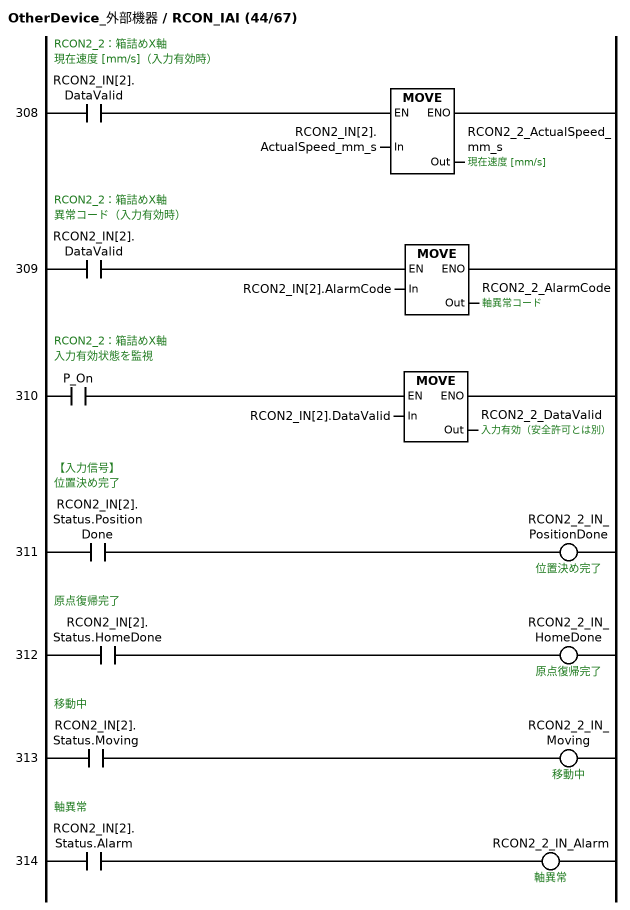
(* [picture p120: OtherDevice_外部機器 / RCON_IAI, rungs 308-314] *)
(* Rung 308: RCON2_2：箱詰めX軸 / 現在速度 [mm/s]（入力有効時） *)
IF RCON2_IN[2].DataValid THEN RCON2_2_ActualSpeed_mm_s := RCON2_IN[2].ActualSpeed_mm_s; END_IF;
(* Rung 309: RCON2_2：箱詰めX軸 / 異常コード（入力有効時） *)
IF RCON2_IN[2].DataValid THEN RCON2_2_AlarmCode := RCON2_IN[2].AlarmCode; END_IF;
(* Rung 310: RCON2_2：箱詰めX軸 / 入力有効状態を監視 *)
IF P_On THEN RCON2_2_DataValid := RCON2_IN[2].DataValid; END_IF;
(* Rung 311: 【入力信号】 / 位置決め完了 *)
RCON2_2_IN_PositionDone := RCON2_IN[2].Status.PositionDone;
(* Rung 312: 原点復帰完了 *)
RCON2_2_IN_HomeDone := RCON2_IN[2].Status.HomeDone;
(* Rung 313: 移動中 *)
RCON2_2_IN_Moving := RCON2_IN[2].Status.Moving;
(* Rung 314: 軸異常 *)
RCON2_2_IN_Alarm := RCON2_IN[2].Status.Alarm;

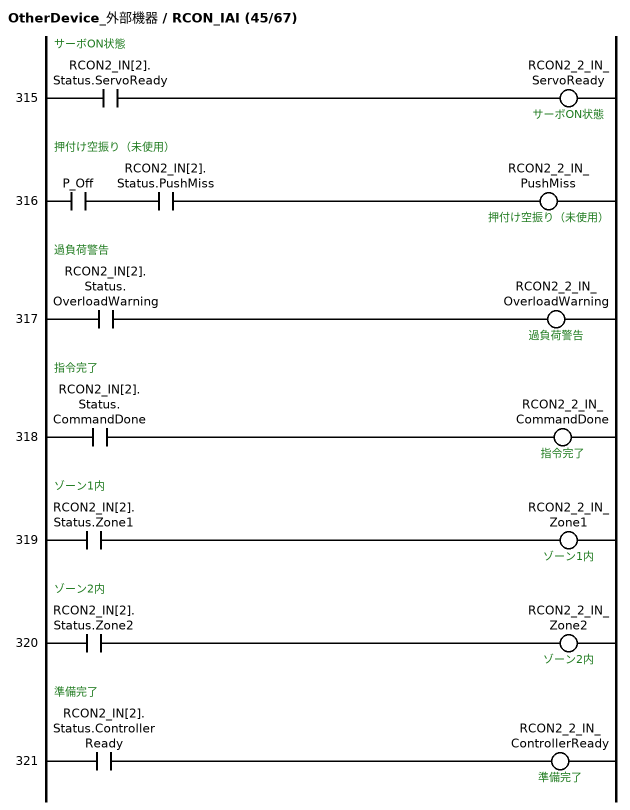
(* Rung 315: サーボON状態 *)
RCON2_2_IN_ServoReady := RCON2_IN[2].Status.ServoReady;
(* Rung 316: 押付け空振り（未使用） *)
RCON2_2_IN_PushMiss := P_Off AND RCON2_IN[2].Status.PushMiss;
(* Rung 317: 過負荷警告 *)
RCON2_2_IN_OverloadWarning := RCON2_IN[2].Status.OverloadWarning;
(* Rung 318: 指令完了 *)
RCON2_2_IN_CommandDone := RCON2_IN[2].Status.CommandDone;
(* Rung 319: ゾーン1内 *)
RCON2_2_IN_Zone1 := RCON2_IN[2].Status.Zone1;
(* Rung 320: ゾーン2内 *)
RCON2_2_IN_Zone2 := RCON2_IN[2].Status.Zone2;
(* Rung 321: 準備完了 *)
RCON2_2_IN_ControllerReady := RCON2_IN[2].Status.ControllerReady;

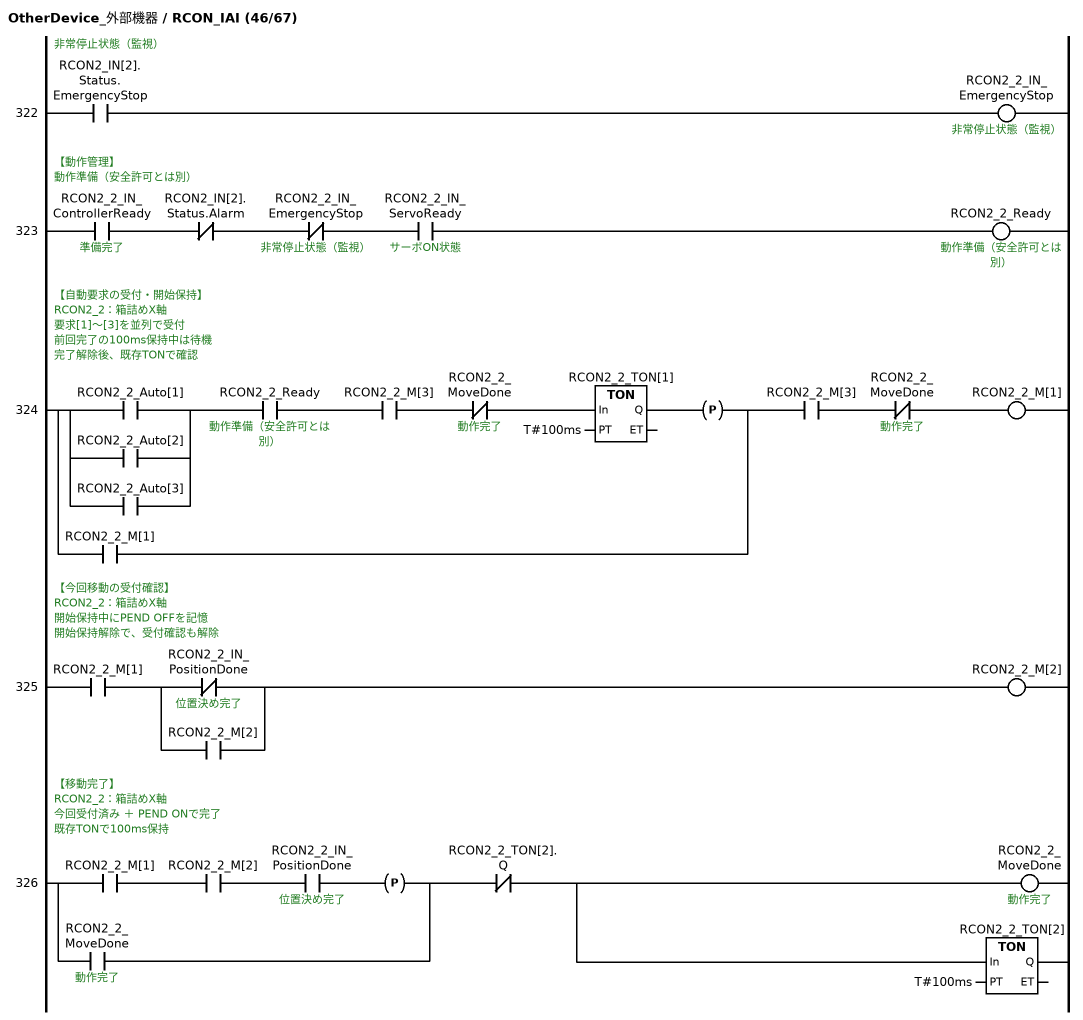
(* Rung 322: 非常停止状態（監視） *)
RCON2_2_IN_EmergencyStop := RCON2_IN[2].Status.EmergencyStop;
(* Rung 323: 【動作管理】 / 動作準備（安全許可とは別） *)
RCON2_2_Ready := RCON2_2_IN_ControllerReady AND NOT RCON2_IN[2].Status.Alarm AND NOT RCON2_2_IN_EmergencyStop AND RCON2_2_IN_ServoReady;
(* Rung 324: 【自動要求の受付・開始保持】 / RCON2_2：箱詰めX軸 / 要求[1]～[3]を並列で受付 / 前回完了の100ms保持中は待機 / 完了解除後、既存TONで確認 *)
RCON2_2_TON[1](In := (RCON2_2_Auto[1] OR RCON2_2_Auto[2] OR RCON2_2_Auto[3]) AND RCON2_2_Ready AND RCON2_2_M[3] AND NOT RCON2_2_MoveDone, PT := T#100ms);
_e30(CLK := RCON2_2_TON[1].Q);
RCON2_2_M[1] := (_e30.Q OR RCON2_2_M[1]) AND RCON2_2_M[3] AND NOT RCON2_2_MoveDone;
(* Rung 325: 【今回移動の受付確認】 / RCON2_2：箱詰めX軸 / 開始保持中にPEND OFFを記憶 / 開始保持解除で、受付確認も解除 *)
RCON2_2_M[2] := RCON2_2_M[1] AND (NOT RCON2_2_IN_PositionDone OR RCON2_2_M[2]);
(* Rung 326: 【移動完了】 / RCON2_2：箱詰めX軸 / 今回受付済み ＋ PEND ONで完了 / 既存TONで100ms保持 *)
_e31(CLK := RCON2_2_M[1] AND RCON2_2_M[2] AND RCON2_2_IN_PositionDone);
_p32 := (_e31.Q OR RCON2_2_MoveDone) AND NOT RCON2_2_TON[2].Q;
RCON2_2_MoveDone := _p32;
RCON2_2_TON[2](In := _p32, PT := T#100ms);

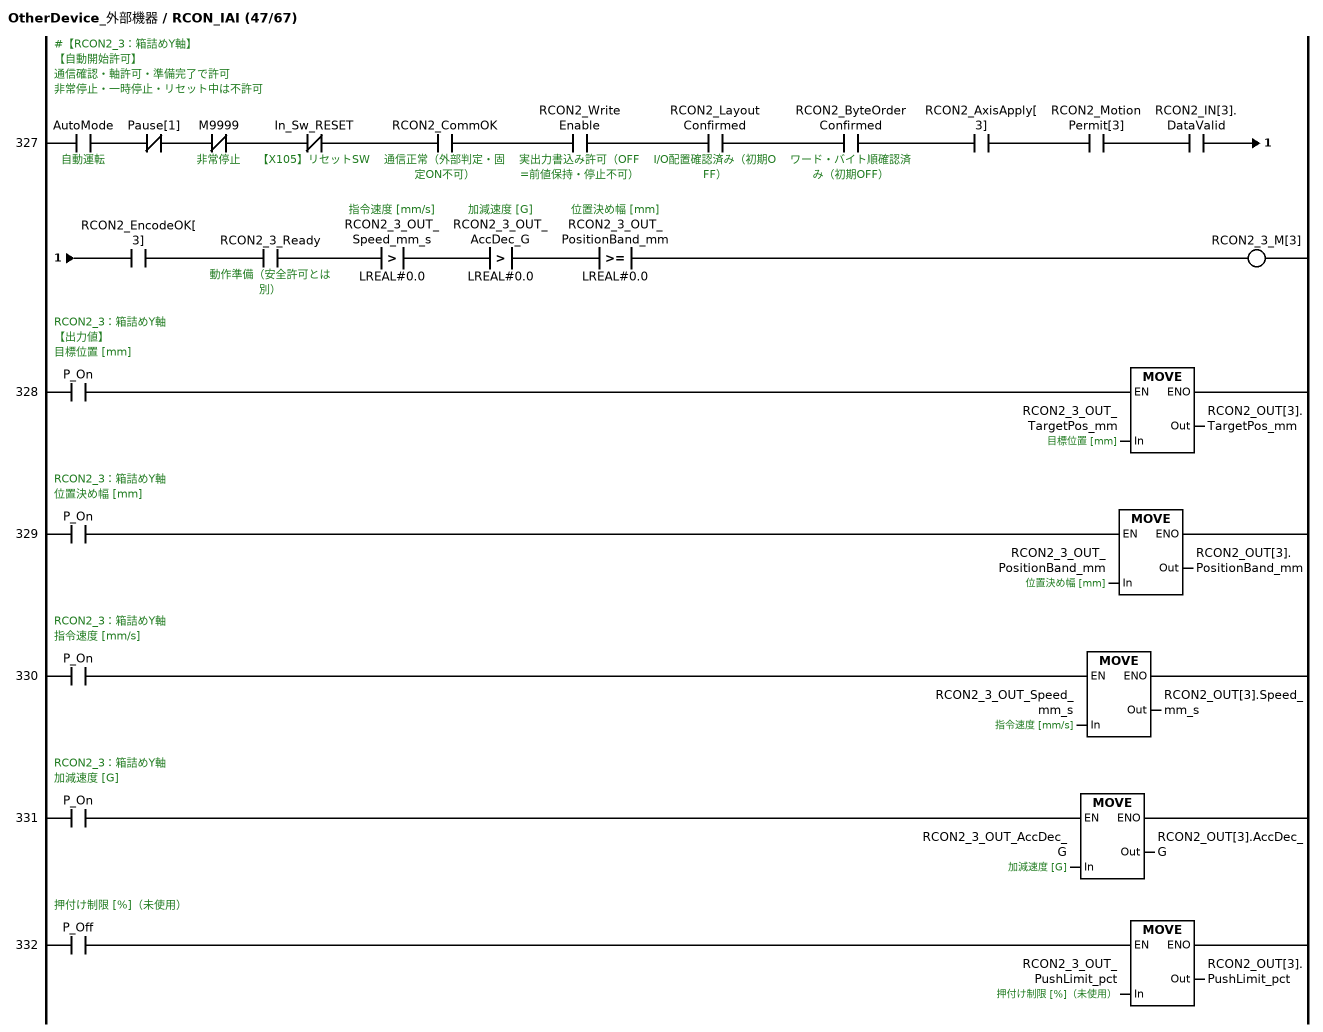
(* Rung 327: #【RCON2_3：箱詰めY軸】 / 【自動開始許可】 / 通信確認・軸許可・準備完了で許可 / 非常停止・一時停止・リセット中は不許可 *)
RCON2_3_M[3] := AutoMode AND NOT Pause[1] AND NOT M9999 AND NOT In_Sw_RESET AND RCON2_CommOK AND RCON2_WriteEnable AND RCON2_LayoutConfirmed AND RCON2_ByteOrderConfirmed AND RCON2_AxisApply[3] AND RCON2_MotionPermit[3] AND RCON2_IN[3].DataValid AND RCON2_EncodeOK[3] AND RCON2_3_Ready AND (RCON2_3_OUT_Speed_mm_s > LREAL#0.0) AND (RCON2_3_OUT_AccDec_G > LREAL#0.0) AND (RCON2_3_OUT_PositionBand_mm >= LREAL#0.0);
(* Rung 328: RCON2_3：箱詰めY軸 / 【出力値】 / 目標位置 [mm] *)
IF P_On THEN RCON2_OUT[3].TargetPos_mm := RCON2_3_OUT_TargetPos_mm; END_IF;
(* Rung 329: RCON2_3：箱詰めY軸 / 位置決め幅 [mm] *)
IF P_On THEN RCON2_OUT[3].PositionBand_mm := RCON2_3_OUT_PositionBand_mm; END_IF;
(* Rung 330: RCON2_3：箱詰めY軸 / 指令速度 [mm/s] *)
IF P_On THEN RCON2_OUT[3].Speed_mm_s := RCON2_3_OUT_Speed_mm_s; END_IF;
(* Rung 331: RCON2_3：箱詰めY軸 / 加減速度 [G] *)
IF P_On THEN RCON2_OUT[3].AccDec_G := RCON2_3_OUT_AccDec_G; END_IF;
(* Rung 332: 押付け制限 [%]（未使用） *)
IF P_Off THEN RCON2_OUT[3].PushLimit_pct := RCON2_3_OUT_PushLimit_pct; END_IF;

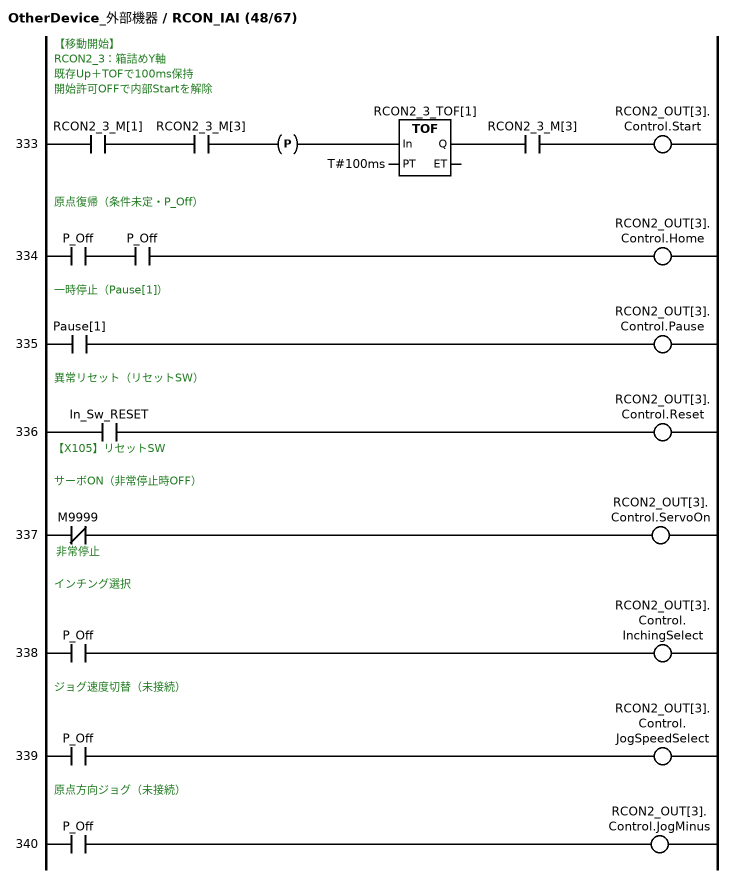
(* Rung 333: 【移動開始】 / RCON2_3：箱詰めY軸 / 既存Up＋TOFで100ms保持 / 開始許可OFFで内部Startを解除 *)
_e33(CLK := RCON2_3_M[1] AND RCON2_3_M[3]);
RCON2_3_TOF[1](In := _e33.Q, PT := T#100ms);
RCON2_OUT[3].Control.Start := RCON2_3_TOF[1].Q AND RCON2_3_M[3];
(* Rung 334: 原点復帰（条件未定・P_Off） *)
RCON2_OUT[3].Control.Home := P_Off AND P_Off;
(* Rung 335: 一時停止（Pause[1]） *)
RCON2_OUT[3].Control.Pause := Pause[1];
(* Rung 336: 異常リセット（リセットSW） *)
RCON2_OUT[3].Control.Reset := In_Sw_RESET;
(* Rung 337: サーボON（非常停止時OFF） *)
RCON2_OUT[3].Control.ServoOn := NOT M9999;
(* Rung 338: インチング選択 *)
RCON2_OUT[3].Control.InchingSelect := P_Off;
(* Rung 339: ジョグ速度切替（未接続） *)
RCON2_OUT[3].Control.JogSpeedSelect := P_Off;
(* Rung 340: 原点方向ジョグ（未接続） *)
RCON2_OUT[3].Control.JogMinus := P_Off;

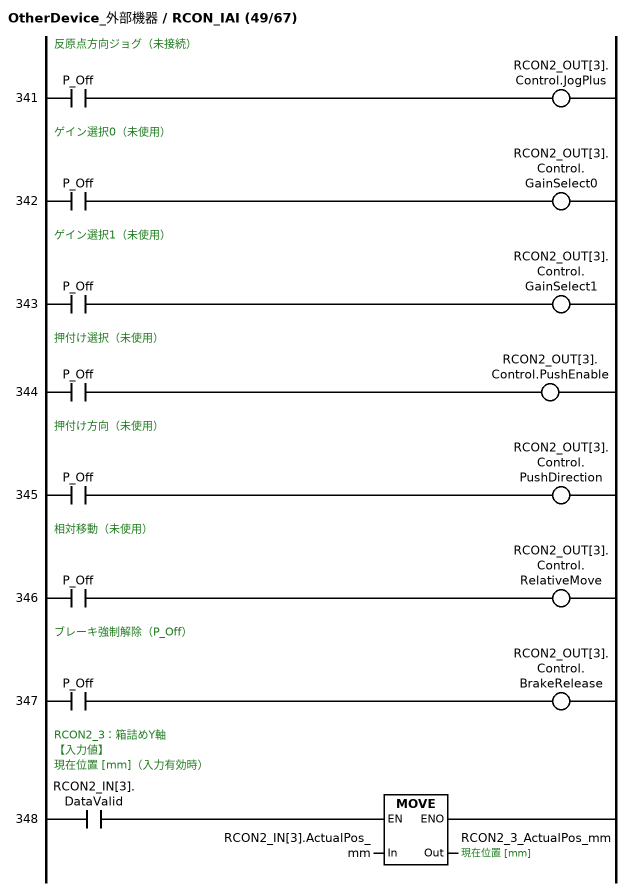
(* Rung 341: 反原点方向ジョグ（未接続） *)
RCON2_OUT[3].Control.JogPlus := P_Off;
(* Rung 342: ゲイン選択0（未使用） *)
RCON2_OUT[3].Control.GainSelect0 := P_Off;
(* Rung 343: ゲイン選択1（未使用） *)
RCON2_OUT[3].Control.GainSelect1 := P_Off;
(* Rung 344: 押付け選択（未使用） *)
RCON2_OUT[3].Control.PushEnable := P_Off;
(* Rung 345: 押付け方向（未使用） *)
RCON2_OUT[3].Control.PushDirection := P_Off;
(* Rung 346: 相対移動（未使用） *)
RCON2_OUT[3].Control.RelativeMove := P_Off;
(* Rung 347: ブレーキ強制解除（P_Off） *)
RCON2_OUT[3].Control.BrakeRelease := P_Off;
(* Rung 348: RCON2_3：箱詰めY軸 / 【入力値】 / 現在位置 [mm]（入力有効時） *)
IF RCON2_IN[3].DataValid THEN RCON2_3_ActualPos_mm := RCON2_IN[3].ActualPos_mm; END_IF;

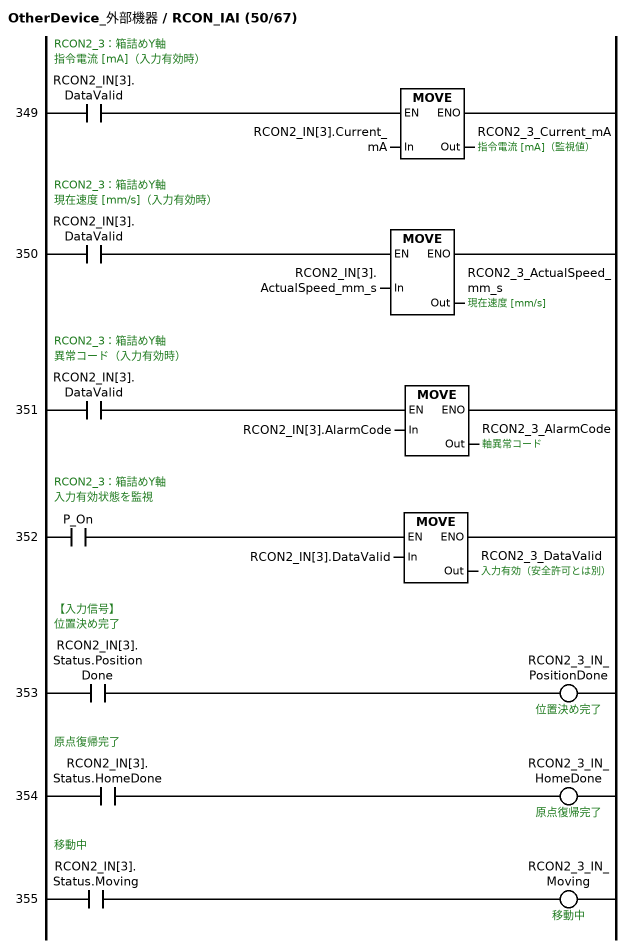
(* Rung 349: RCON2_3：箱詰めY軸 / 指令電流 [mA]（入力有効時） *)
IF RCON2_IN[3].DataValid THEN RCON2_3_Current_mA := RCON2_IN[3].Current_mA; END_IF;
(* Rung 350: RCON2_3：箱詰めY軸 / 現在速度 [mm/s]（入力有効時） *)
IF RCON2_IN[3].DataValid THEN RCON2_3_ActualSpeed_mm_s := RCON2_IN[3].ActualSpeed_mm_s; END_IF;
(* Rung 351: RCON2_3：箱詰めY軸 / 異常コード（入力有効時） *)
IF RCON2_IN[3].DataValid THEN RCON2_3_AlarmCode := RCON2_IN[3].AlarmCode; END_IF;
(* Rung 352: RCON2_3：箱詰めY軸 / 入力有効状態を監視 *)
IF P_On THEN RCON2_3_DataValid := RCON2_IN[3].DataValid; END_IF;
(* Rung 353: 【入力信号】 / 位置決め完了 *)
RCON2_3_IN_PositionDone := RCON2_IN[3].Status.PositionDone;
(* Rung 354: 原点復帰完了 *)
RCON2_3_IN_HomeDone := RCON2_IN[3].Status.HomeDone;
(* Rung 355: 移動中 *)
RCON2_3_IN_Moving := RCON2_IN[3].Status.Moving;

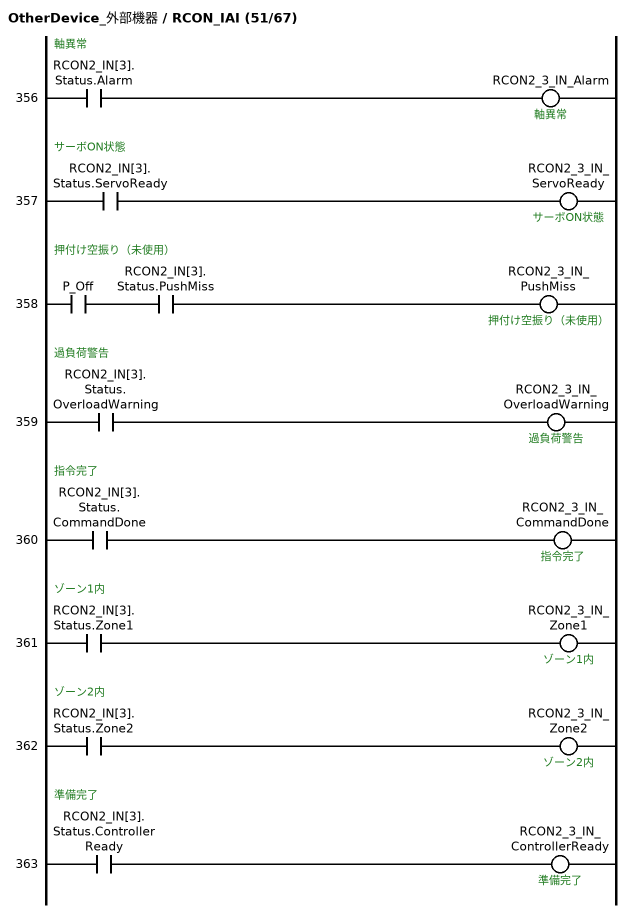
(* Rung 356: 軸異常 *)
RCON2_3_IN_Alarm := RCON2_IN[3].Status.Alarm;
(* Rung 357: サーボON状態 *)
RCON2_3_IN_ServoReady := RCON2_IN[3].Status.ServoReady;
(* Rung 358: 押付け空振り（未使用） *)
RCON2_3_IN_PushMiss := P_Off AND RCON2_IN[3].Status.PushMiss;
(* Rung 359: 過負荷警告 *)
RCON2_3_IN_OverloadWarning := RCON2_IN[3].Status.OverloadWarning;
(* Rung 360: 指令完了 *)
RCON2_3_IN_CommandDone := RCON2_IN[3].Status.CommandDone;
(* Rung 361: ゾーン1内 *)
RCON2_3_IN_Zone1 := RCON2_IN[3].Status.Zone1;
(* Rung 362: ゾーン2内 *)
RCON2_3_IN_Zone2 := RCON2_IN[3].Status.Zone2;
(* Rung 363: 準備完了 *)
RCON2_3_IN_ControllerReady := RCON2_IN[3].Status.ControllerReady;

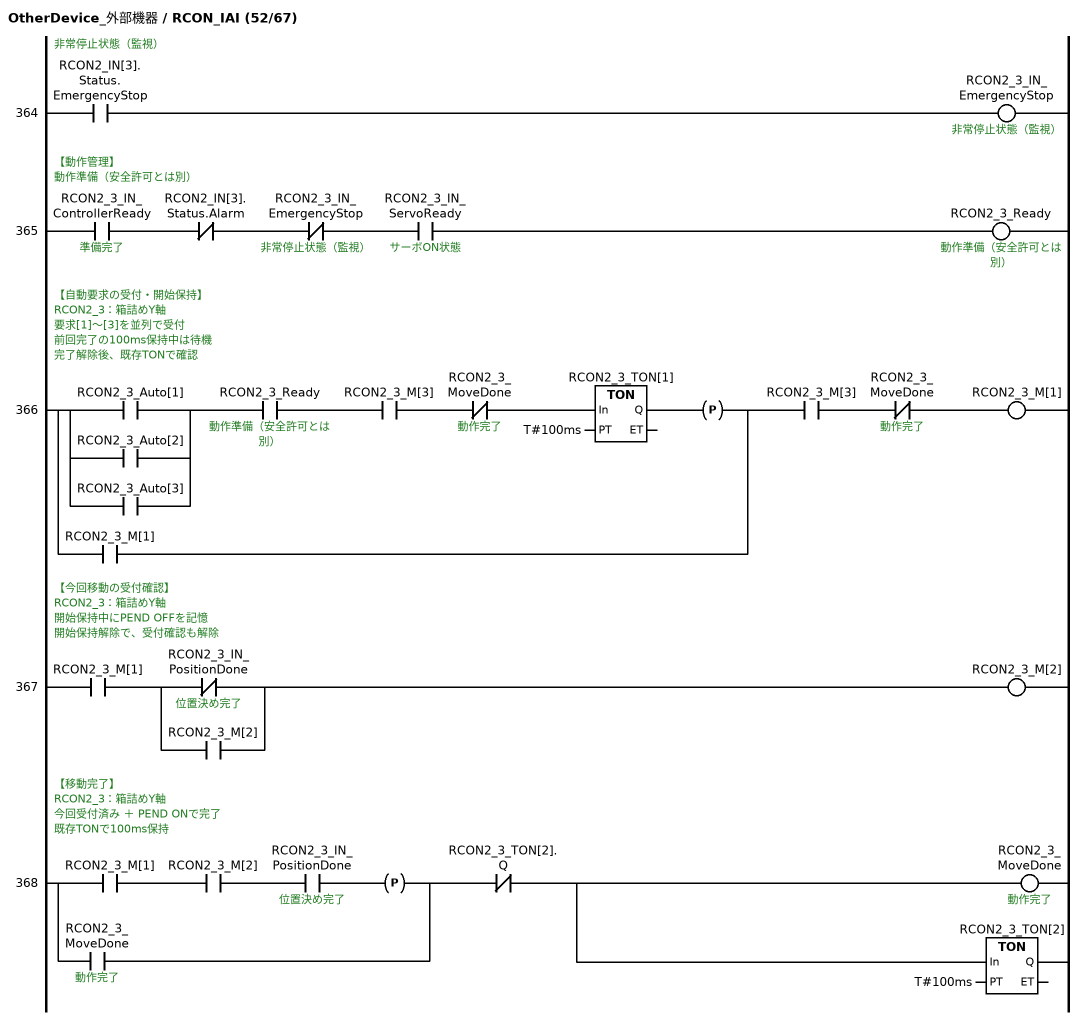
(* Rung 364: 非常停止状態（監視） *)
RCON2_3_IN_EmergencyStop := RCON2_IN[3].Status.EmergencyStop;
(* Rung 365: 【動作管理】 / 動作準備（安全許可とは別） *)
RCON2_3_Ready := RCON2_3_IN_ControllerReady AND NOT RCON2_IN[3].Status.Alarm AND NOT RCON2_3_IN_EmergencyStop AND RCON2_3_IN_ServoReady;
(* Rung 366: 【自動要求の受付・開始保持】 / RCON2_3：箱詰めY軸 / 要求[1]～[3]を並列で受付 / 前回完了の100ms保持中は待機 / 完了解除後、既存TONで確認 *)
RCON2_3_TON[1](In := (RCON2_3_Auto[1] OR RCON2_3_Auto[2] OR RCON2_3_Auto[3]) AND RCON2_3_Ready AND RCON2_3_M[3] AND NOT RCON2_3_MoveDone, PT := T#100ms);
_e34(CLK := RCON2_3_TON[1].Q);
RCON2_3_M[1] := (_e34.Q OR RCON2_3_M[1]) AND RCON2_3_M[3] AND NOT RCON2_3_MoveDone;
(* Rung 367: 【今回移動の受付確認】 / RCON2_3：箱詰めY軸 / 開始保持中にPEND OFFを記憶 / 開始保持解除で、受付確認も解除 *)
RCON2_3_M[2] := RCON2_3_M[1] AND (NOT RCON2_3_IN_PositionDone OR RCON2_3_M[2]);
(* Rung 368: 【移動完了】 / RCON2_3：箱詰めY軸 / 今回受付済み ＋ PEND ONで完了 / 既存TONで100ms保持 *)
_e35(CLK := RCON2_3_M[1] AND RCON2_3_M[2] AND RCON2_3_IN_PositionDone);
_p36 := (_e35.Q OR RCON2_3_MoveDone) AND NOT RCON2_3_TON[2].Q;
RCON2_3_MoveDone := _p36;
RCON2_3_TON[2](In := _p36, PT := T#100ms);

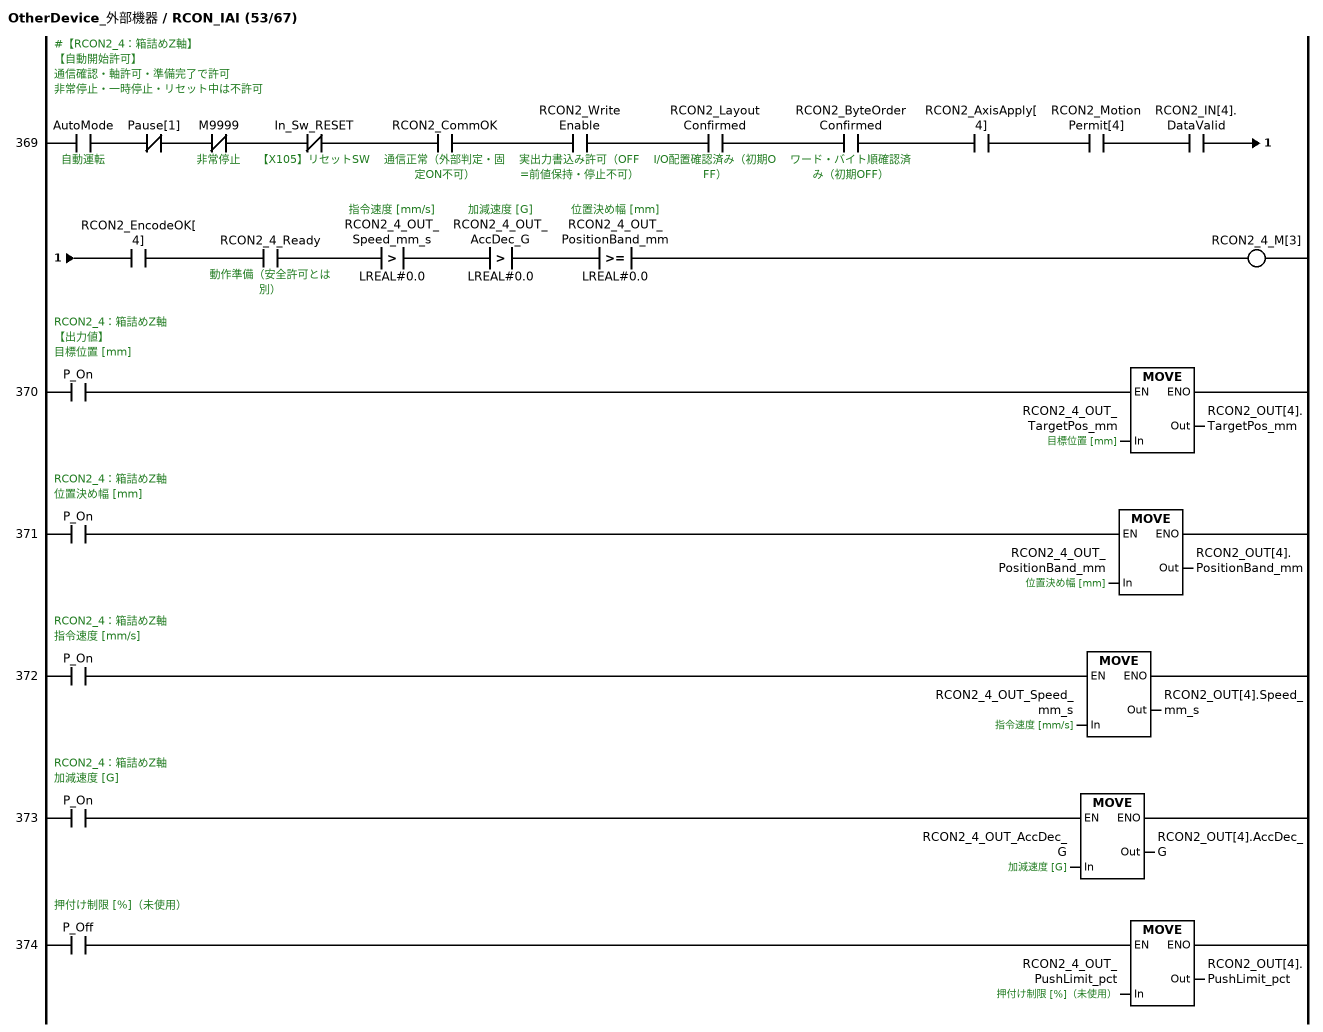
(* Rung 369: #【RCON2_4：箱詰めZ軸】 / 【自動開始許可】 / 通信確認・軸許可・準備完了で許可 / 非常停止・一時停止・リセット中は不許可 *)
RCON2_4_M[3] := AutoMode AND NOT Pause[1] AND NOT M9999 AND NOT In_Sw_RESET AND RCON2_CommOK AND RCON2_WriteEnable AND RCON2_LayoutConfirmed AND RCON2_ByteOrderConfirmed AND RCON2_AxisApply[4] AND RCON2_MotionPermit[4] AND RCON2_IN[4].DataValid AND RCON2_EncodeOK[4] AND RCON2_4_Ready AND (RCON2_4_OUT_Speed_mm_s > LREAL#0.0) AND (RCON2_4_OUT_AccDec_G > LREAL#0.0) AND (RCON2_4_OUT_PositionBand_mm >= LREAL#0.0);
(* Rung 370: RCON2_4：箱詰めZ軸 / 【出力値】 / 目標位置 [mm] *)
IF P_On THEN RCON2_OUT[4].TargetPos_mm := RCON2_4_OUT_TargetPos_mm; END_IF;
(* Rung 371: RCON2_4：箱詰めZ軸 / 位置決め幅 [mm] *)
IF P_On THEN RCON2_OUT[4].PositionBand_mm := RCON2_4_OUT_PositionBand_mm; END_IF;
(* Rung 372: RCON2_4：箱詰めZ軸 / 指令速度 [mm/s] *)
IF P_On THEN RCON2_OUT[4].Speed_mm_s := RCON2_4_OUT_Speed_mm_s; END_IF;
(* Rung 373: RCON2_4：箱詰めZ軸 / 加減速度 [G] *)
IF P_On THEN RCON2_OUT[4].AccDec_G := RCON2_4_OUT_AccDec_G; END_IF;
(* Rung 374: 押付け制限 [%]（未使用） *)
IF P_Off THEN RCON2_OUT[4].PushLimit_pct := RCON2_4_OUT_PushLimit_pct; END_IF;

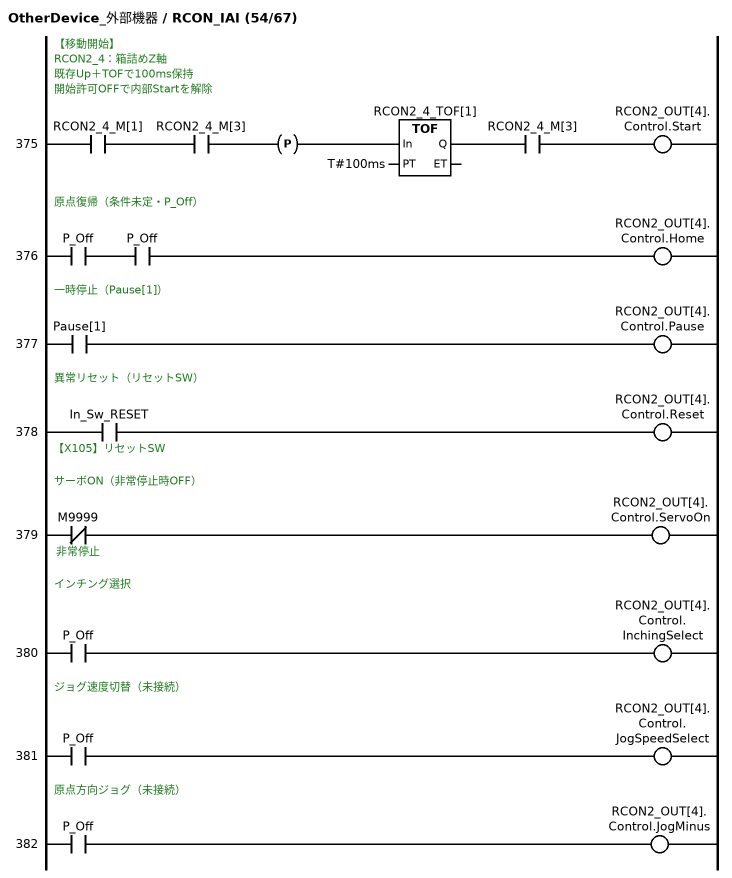
(* Rung 375: 【移動開始】 / RCON2_4：箱詰めZ軸 / 既存Up＋TOFで100ms保持 / 開始許可OFFで内部Startを解除 *)
_e37(CLK := RCON2_4_M[1] AND RCON2_4_M[3]);
RCON2_4_TOF[1](In := _e37.Q, PT := T#100ms);
RCON2_OUT[4].Control.Start := RCON2_4_TOF[1].Q AND RCON2_4_M[3];
(* Rung 376: 原点復帰（条件未定・P_Off） *)
RCON2_OUT[4].Control.Home := P_Off AND P_Off;
(* Rung 377: 一時停止（Pause[1]） *)
RCON2_OUT[4].Control.Pause := Pause[1];
(* Rung 378: 異常リセット（リセットSW） *)
RCON2_OUT[4].Control.Reset := In_Sw_RESET;
(* Rung 379: サーボON（非常停止時OFF） *)
RCON2_OUT[4].Control.ServoOn := NOT M9999;
(* Rung 380: インチング選択 *)
RCON2_OUT[4].Control.InchingSelect := P_Off;
(* Rung 381: ジョグ速度切替（未接続） *)
RCON2_OUT[4].Control.JogSpeedSelect := P_Off;
(* Rung 382: 原点方向ジョグ（未接続） *)
RCON2_OUT[4].Control.JogMinus := P_Off;

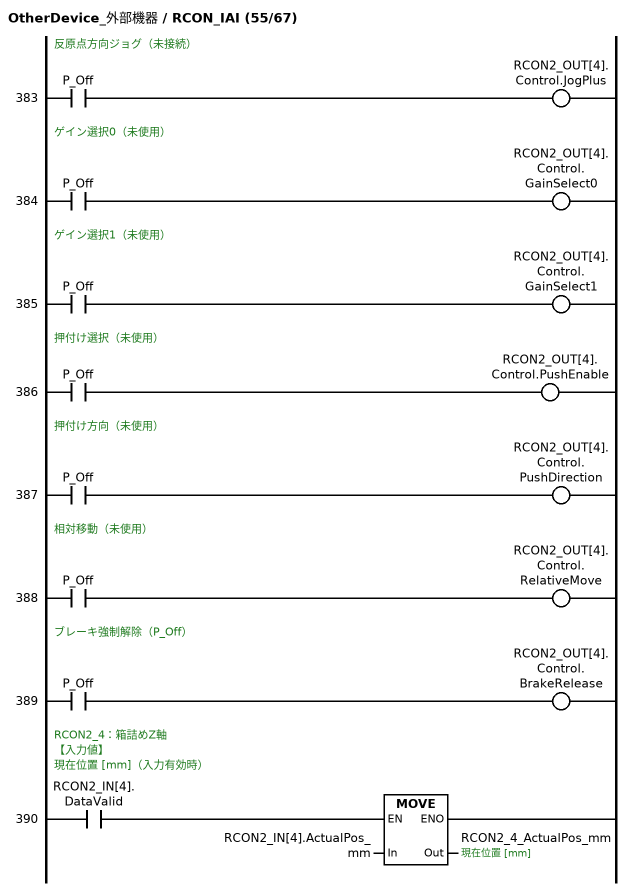
(* Rung 383: 反原点方向ジョグ（未接続） *)
RCON2_OUT[4].Control.JogPlus := P_Off;
(* Rung 384: ゲイン選択0（未使用） *)
RCON2_OUT[4].Control.GainSelect0 := P_Off;
(* Rung 385: ゲイン選択1（未使用） *)
RCON2_OUT[4].Control.GainSelect1 := P_Off;
(* Rung 386: 押付け選択（未使用） *)
RCON2_OUT[4].Control.PushEnable := P_Off;
(* Rung 387: 押付け方向（未使用） *)
RCON2_OUT[4].Control.PushDirection := P_Off;
(* Rung 388: 相対移動（未使用） *)
RCON2_OUT[4].Control.RelativeMove := P_Off;
(* Rung 389: ブレーキ強制解除（P_Off） *)
RCON2_OUT[4].Control.BrakeRelease := P_Off;
(* Rung 390: RCON2_4：箱詰めZ軸 / 【入力値】 / 現在位置 [mm]（入力有効時） *)
IF RCON2_IN[4].DataValid THEN RCON2_4_ActualPos_mm := RCON2_IN[4].ActualPos_mm; END_IF;

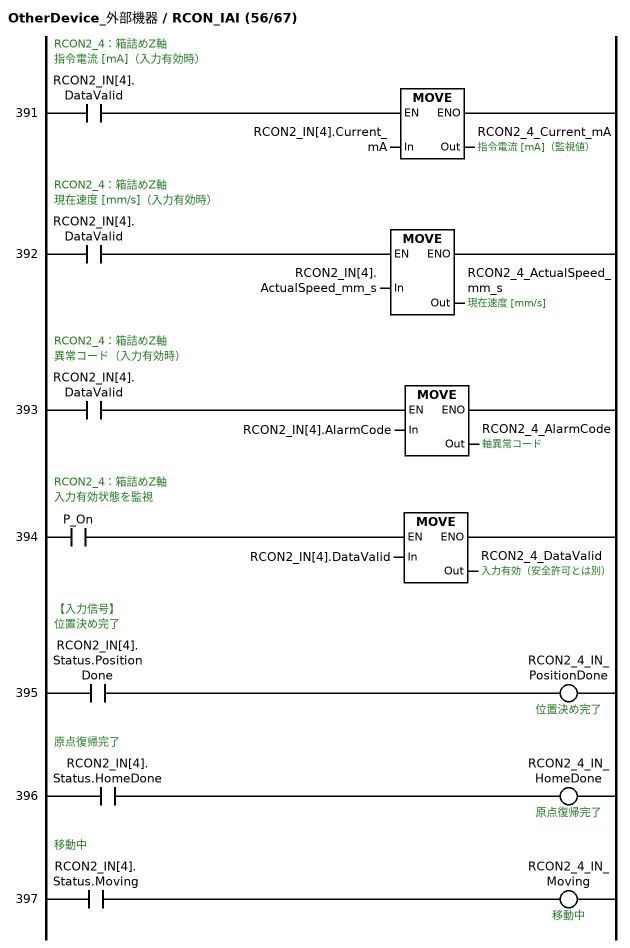
(* Rung 391: RCON2_4：箱詰めZ軸 / 指令電流 [mA]（入力有効時） *)
IF RCON2_IN[4].DataValid THEN RCON2_4_Current_mA := RCON2_IN[4].Current_mA; END_IF;
(* Rung 392: RCON2_4：箱詰めZ軸 / 現在速度 [mm/s]（入力有効時） *)
IF RCON2_IN[4].DataValid THEN RCON2_4_ActualSpeed_mm_s := RCON2_IN[4].ActualSpeed_mm_s; END_IF;
(* Rung 393: RCON2_4：箱詰めZ軸 / 異常コード（入力有効時） *)
IF RCON2_IN[4].DataValid THEN RCON2_4_AlarmCode := RCON2_IN[4].AlarmCode; END_IF;
(* Rung 394: RCON2_4：箱詰めZ軸 / 入力有効状態を監視 *)
IF P_On THEN RCON2_4_DataValid := RCON2_IN[4].DataValid; END_IF;
(* Rung 395: 【入力信号】 / 位置決め完了 *)
RCON2_4_IN_PositionDone := RCON2_IN[4].Status.PositionDone;
(* Rung 396: 原点復帰完了 *)
RCON2_4_IN_HomeDone := RCON2_IN[4].Status.HomeDone;
(* Rung 397: 移動中 *)
RCON2_4_IN_Moving := RCON2_IN[4].Status.Moving;

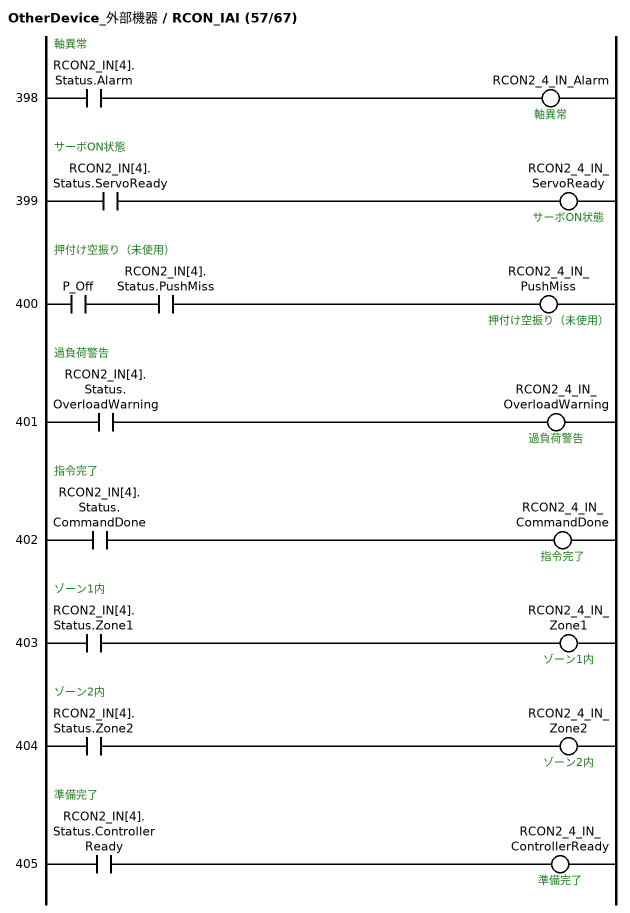
(* Rung 398: 軸異常 *)
RCON2_4_IN_Alarm := RCON2_IN[4].Status.Alarm;
(* Rung 399: サーボON状態 *)
RCON2_4_IN_ServoReady := RCON2_IN[4].Status.ServoReady;
(* Rung 400: 押付け空振り（未使用） *)
RCON2_4_IN_PushMiss := P_Off AND RCON2_IN[4].Status.PushMiss;
(* Rung 401: 過負荷警告 *)
RCON2_4_IN_OverloadWarning := RCON2_IN[4].Status.OverloadWarning;
(* Rung 402: 指令完了 *)
RCON2_4_IN_CommandDone := RCON2_IN[4].Status.CommandDone;
(* Rung 403: ゾーン1内 *)
RCON2_4_IN_Zone1 := RCON2_IN[4].Status.Zone1;
(* Rung 404: ゾーン2内 *)
RCON2_4_IN_Zone2 := RCON2_IN[4].Status.Zone2;
(* Rung 405: 準備完了 *)
RCON2_4_IN_ControllerReady := RCON2_IN[4].Status.ControllerReady;

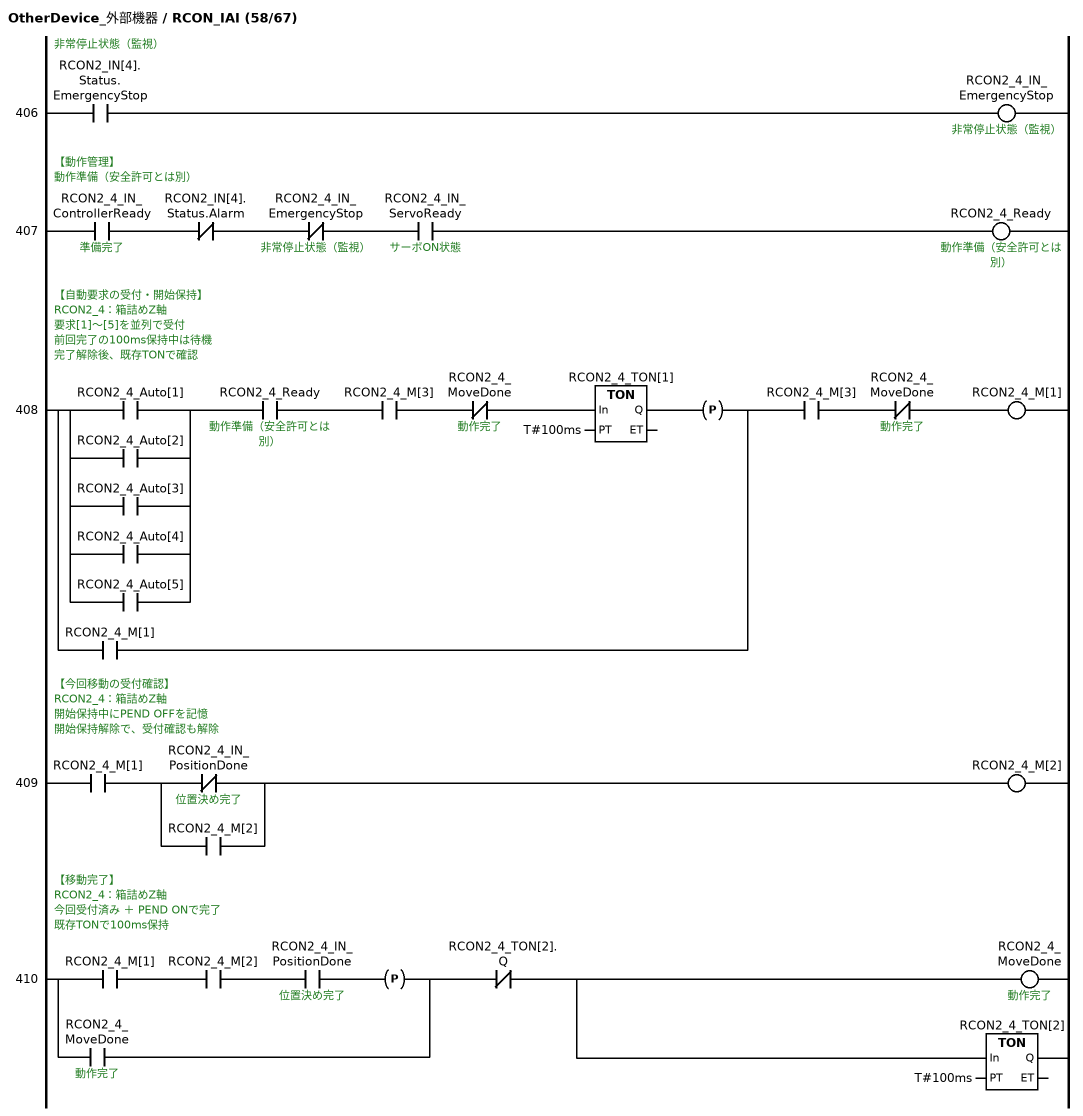
(* Rung 406: 非常停止状態（監視） *)
RCON2_4_IN_EmergencyStop := RCON2_IN[4].Status.EmergencyStop;
(* Rung 407: 【動作管理】 / 動作準備（安全許可とは別） *)
RCON2_4_Ready := RCON2_4_IN_ControllerReady AND NOT RCON2_IN[4].Status.Alarm AND NOT RCON2_4_IN_EmergencyStop AND RCON2_4_IN_ServoReady;
(* Rung 408: 【自動要求の受付・開始保持】 / RCON2_4：箱詰めZ軸 / 要求[1]～[5]を並列で受付 / 前回完了の100ms保持中は待機 / 完了解除後、既存TONで確認 *)
RCON2_4_TON[1](In := (RCON2_4_Auto[1] OR RCON2_4_Auto[2] OR RCON2_4_Auto[3] OR RCON2_4_Auto[4] OR RCON2_4_Auto[5]) AND RCON2_4_Ready AND RCON2_4_M[3] AND NOT RCON2_4_MoveDone, PT := T#100ms);
_e38(CLK := RCON2_4_TON[1].Q);
RCON2_4_M[1] := (_e38.Q OR RCON2_4_M[1]) AND RCON2_4_M[3] AND NOT RCON2_4_MoveDone;
(* Rung 409: 【今回移動の受付確認】 / RCON2_4：箱詰めZ軸 / 開始保持中にPEND OFFを記憶 / 開始保持解除で、受付確認も解除 *)
RCON2_4_M[2] := RCON2_4_M[1] AND (NOT RCON2_4_IN_PositionDone OR RCON2_4_M[2]);
(* Rung 410: 【移動完了】 / RCON2_4：箱詰めZ軸 / 今回受付済み ＋ PEND ONで完了 / 既存TONで100ms保持 *)
_e39(CLK := RCON2_4_M[1] AND RCON2_4_M[2] AND RCON2_4_IN_PositionDone);
_p40 := (_e39.Q OR RCON2_4_MoveDone) AND NOT RCON2_4_TON[2].Q;
RCON2_4_MoveDone := _p40;
RCON2_4_TON[2](In := _p40, PT := T#100ms);

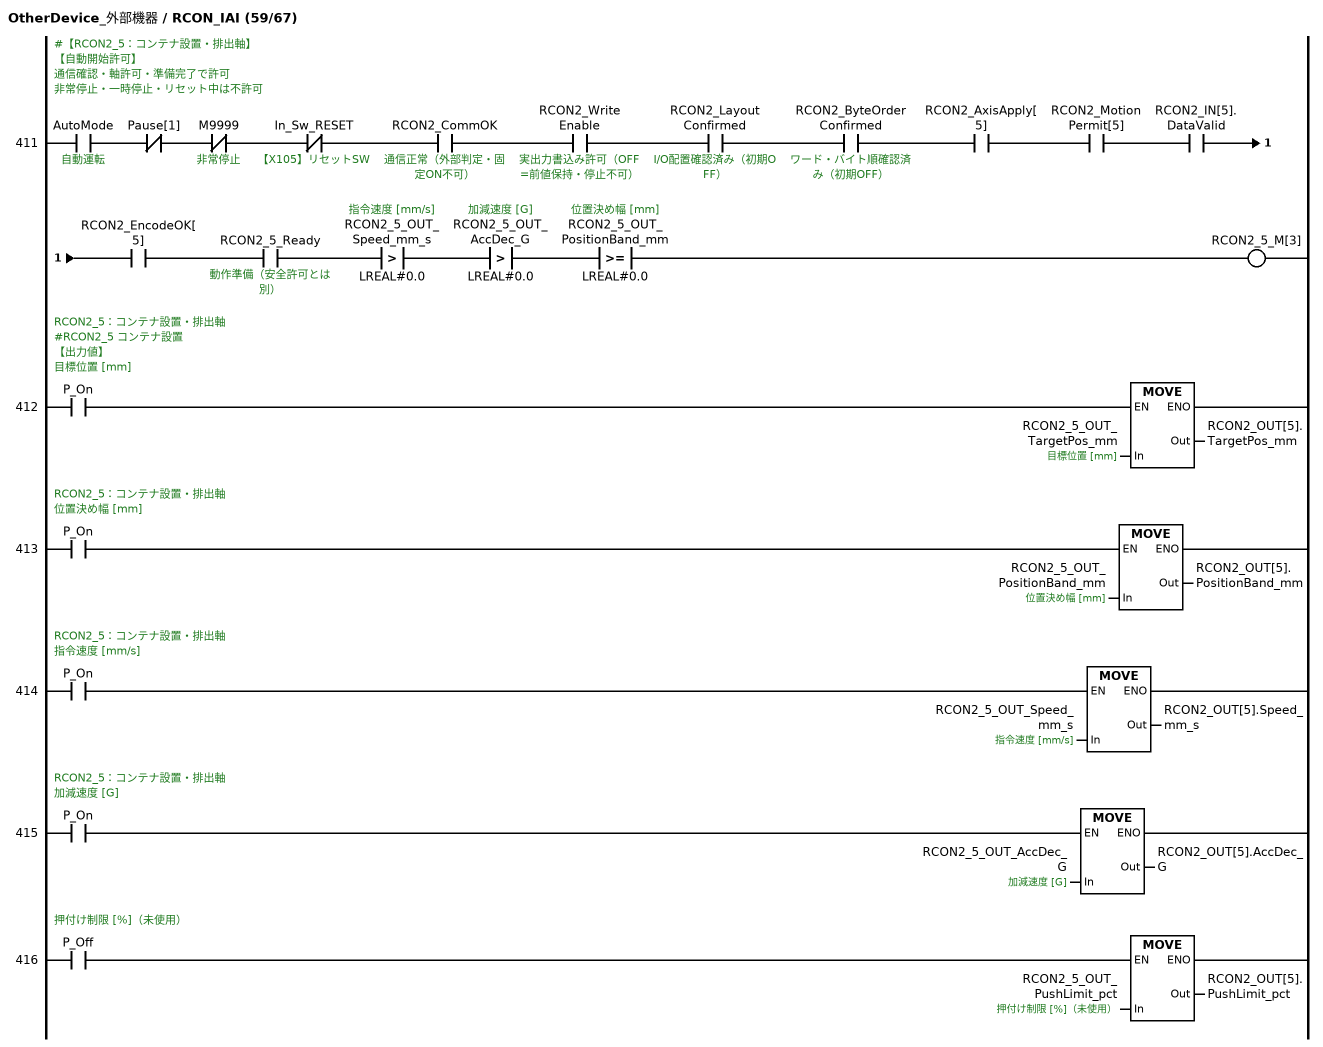
(* Rung 411: #【RCON2_5：コンテナ設置・排出軸】 / 【自動開始許可】 / 通信確認・軸許可・準備完了で許可 / 非常停止・一時停止・リセット中は不許可 *)
RCON2_5_M[3] := AutoMode AND NOT Pause[1] AND NOT M9999 AND NOT In_Sw_RESET AND RCON2_CommOK AND RCON2_WriteEnable AND RCON2_LayoutConfirmed AND RCON2_ByteOrderConfirmed AND RCON2_AxisApply[5] AND RCON2_MotionPermit[5] AND RCON2_IN[5].DataValid AND RCON2_EncodeOK[5] AND RCON2_5_Ready AND (RCON2_5_OUT_Speed_mm_s > LREAL#0.0) AND (RCON2_5_OUT_AccDec_G > LREAL#0.0) AND (RCON2_5_OUT_PositionBand_mm >= LREAL#0.0);
(* Rung 412: RCON2_5：コンテナ設置・排出軸 / #RCON2_5 コンテナ設置 / 【出力値】 / 目標位置 [mm] *)
IF P_On THEN RCON2_OUT[5].TargetPos_mm := RCON2_5_OUT_TargetPos_mm; END_IF;
(* Rung 413: RCON2_5：コンテナ設置・排出軸 / 位置決め幅 [mm] *)
IF P_On THEN RCON2_OUT[5].PositionBand_mm := RCON2_5_OUT_PositionBand_mm; END_IF;
(* Rung 414: RCON2_5：コンテナ設置・排出軸 / 指令速度 [mm/s] *)
IF P_On THEN RCON2_OUT[5].Speed_mm_s := RCON2_5_OUT_Speed_mm_s; END_IF;
(* Rung 415: RCON2_5：コンテナ設置・排出軸 / 加減速度 [G] *)
IF P_On THEN RCON2_OUT[5].AccDec_G := RCON2_5_OUT_AccDec_G; END_IF;
(* Rung 416: 押付け制限 [%]（未使用） *)
IF P_Off THEN RCON2_OUT[5].PushLimit_pct := RCON2_5_OUT_PushLimit_pct; END_IF;

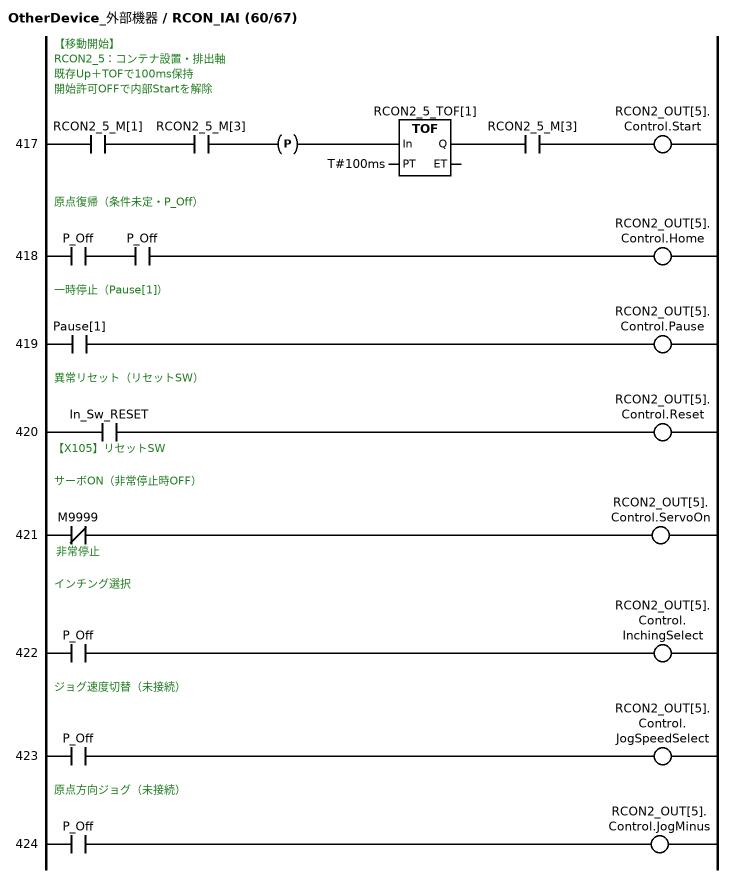
(* Rung 417: 【移動開始】 / RCON2_5：コンテナ設置・排出軸 / 既存Up＋TOFで100ms保持 / 開始許可OFFで内部Startを解除 *)
_e41(CLK := RCON2_5_M[1] AND RCON2_5_M[3]);
RCON2_5_TOF[1](In := _e41.Q, PT := T#100ms);
RCON2_OUT[5].Control.Start := RCON2_5_TOF[1].Q AND RCON2_5_M[3];
(* Rung 418: 原点復帰（条件未定・P_Off） *)
RCON2_OUT[5].Control.Home := P_Off AND P_Off;
(* Rung 419: 一時停止（Pause[1]） *)
RCON2_OUT[5].Control.Pause := Pause[1];
(* Rung 420: 異常リセット（リセットSW） *)
RCON2_OUT[5].Control.Reset := In_Sw_RESET;
(* Rung 421: サーボON（非常停止時OFF） *)
RCON2_OUT[5].Control.ServoOn := NOT M9999;
(* Rung 422: インチング選択 *)
RCON2_OUT[5].Control.InchingSelect := P_Off;
(* Rung 423: ジョグ速度切替（未接続） *)
RCON2_OUT[5].Control.JogSpeedSelect := P_Off;
(* Rung 424: 原点方向ジョグ（未接続） *)
RCON2_OUT[5].Control.JogMinus := P_Off;

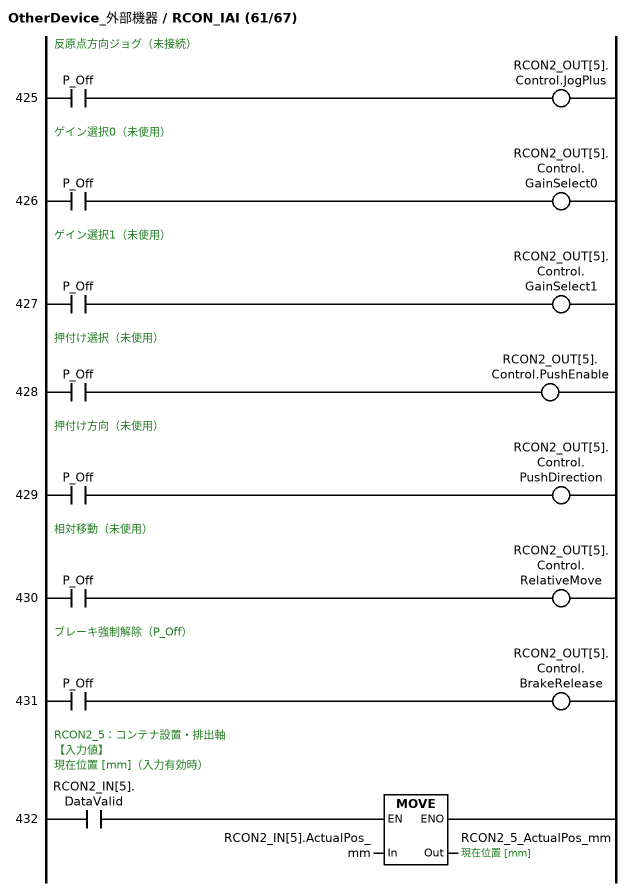
(* Rung 425: 反原点方向ジョグ（未接続） *)
RCON2_OUT[5].Control.JogPlus := P_Off;
(* Rung 426: ゲイン選択0（未使用） *)
RCON2_OUT[5].Control.GainSelect0 := P_Off;
(* Rung 427: ゲイン選択1（未使用） *)
RCON2_OUT[5].Control.GainSelect1 := P_Off;
(* Rung 428: 押付け選択（未使用） *)
RCON2_OUT[5].Control.PushEnable := P_Off;
(* Rung 429: 押付け方向（未使用） *)
RCON2_OUT[5].Control.PushDirection := P_Off;
(* Rung 430: 相対移動（未使用） *)
RCON2_OUT[5].Control.RelativeMove := P_Off;
(* Rung 431: ブレーキ強制解除（P_Off） *)
RCON2_OUT[5].Control.BrakeRelease := P_Off;
(* Rung 432: RCON2_5：コンテナ設置・排出軸 / 【入力値】 / 現在位置 [mm]（入力有効時） *)
IF RCON2_IN[5].DataValid THEN RCON2_5_ActualPos_mm := RCON2_IN[5].ActualPos_mm; END_IF;

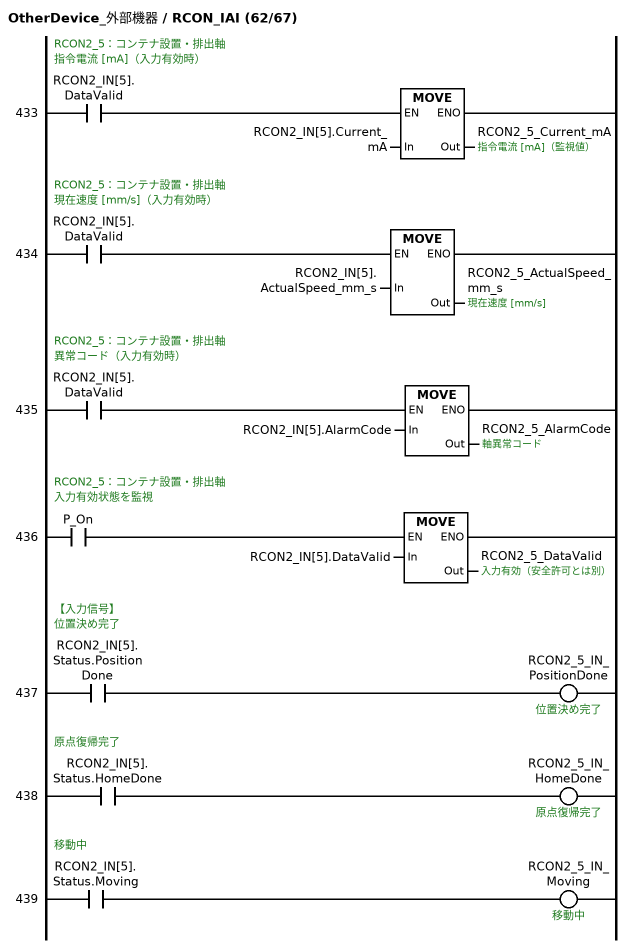
(* Rung 433: RCON2_5：コンテナ設置・排出軸 / 指令電流 [mA]（入力有効時） *)
IF RCON2_IN[5].DataValid THEN RCON2_5_Current_mA := RCON2_IN[5].Current_mA; END_IF;
(* Rung 434: RCON2_5：コンテナ設置・排出軸 / 現在速度 [mm/s]（入力有効時） *)
IF RCON2_IN[5].DataValid THEN RCON2_5_ActualSpeed_mm_s := RCON2_IN[5].ActualSpeed_mm_s; END_IF;
(* Rung 435: RCON2_5：コンテナ設置・排出軸 / 異常コード（入力有効時） *)
IF RCON2_IN[5].DataValid THEN RCON2_5_AlarmCode := RCON2_IN[5].AlarmCode; END_IF;
(* Rung 436: RCON2_5：コンテナ設置・排出軸 / 入力有効状態を監視 *)
IF P_On THEN RCON2_5_DataValid := RCON2_IN[5].DataValid; END_IF;
(* Rung 437: 【入力信号】 / 位置決め完了 *)
RCON2_5_IN_PositionDone := RCON2_IN[5].Status.PositionDone;
(* Rung 438: 原点復帰完了 *)
RCON2_5_IN_HomeDone := RCON2_IN[5].Status.HomeDone;
(* Rung 439: 移動中 *)
RCON2_5_IN_Moving := RCON2_IN[5].Status.Moving;

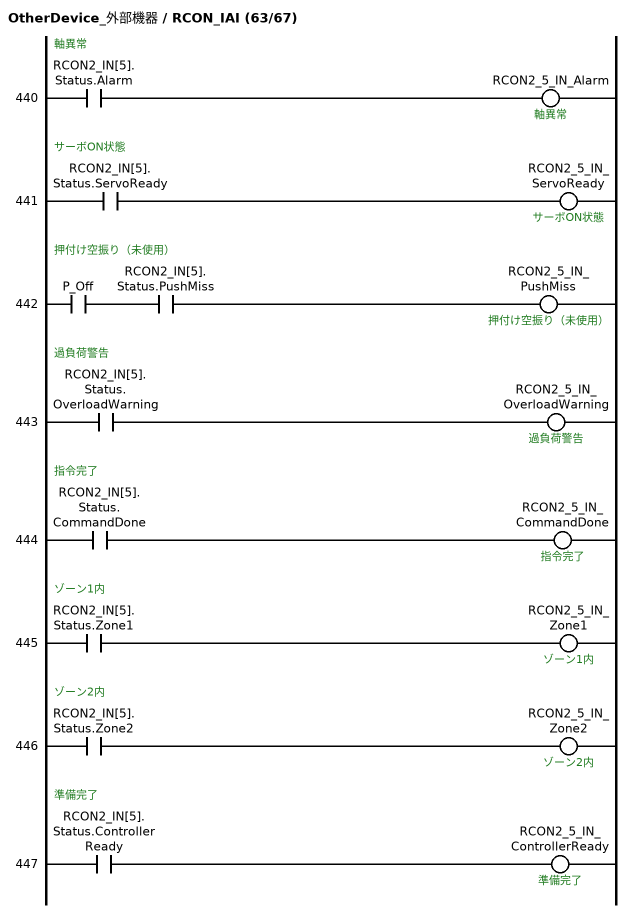
(* Rung 440: 軸異常 *)
RCON2_5_IN_Alarm := RCON2_IN[5].Status.Alarm;
(* Rung 441: サーボON状態 *)
RCON2_5_IN_ServoReady := RCON2_IN[5].Status.ServoReady;
(* Rung 442: 押付け空振り（未使用） *)
RCON2_5_IN_PushMiss := P_Off AND RCON2_IN[5].Status.PushMiss;
(* Rung 443: 過負荷警告 *)
RCON2_5_IN_OverloadWarning := RCON2_IN[5].Status.OverloadWarning;
(* Rung 444: 指令完了 *)
RCON2_5_IN_CommandDone := RCON2_IN[5].Status.CommandDone;
(* Rung 445: ゾーン1内 *)
RCON2_5_IN_Zone1 := RCON2_IN[5].Status.Zone1;
(* Rung 446: ゾーン2内 *)
RCON2_5_IN_Zone2 := RCON2_IN[5].Status.Zone2;
(* Rung 447: 準備完了 *)
RCON2_5_IN_ControllerReady := RCON2_IN[5].Status.ControllerReady;

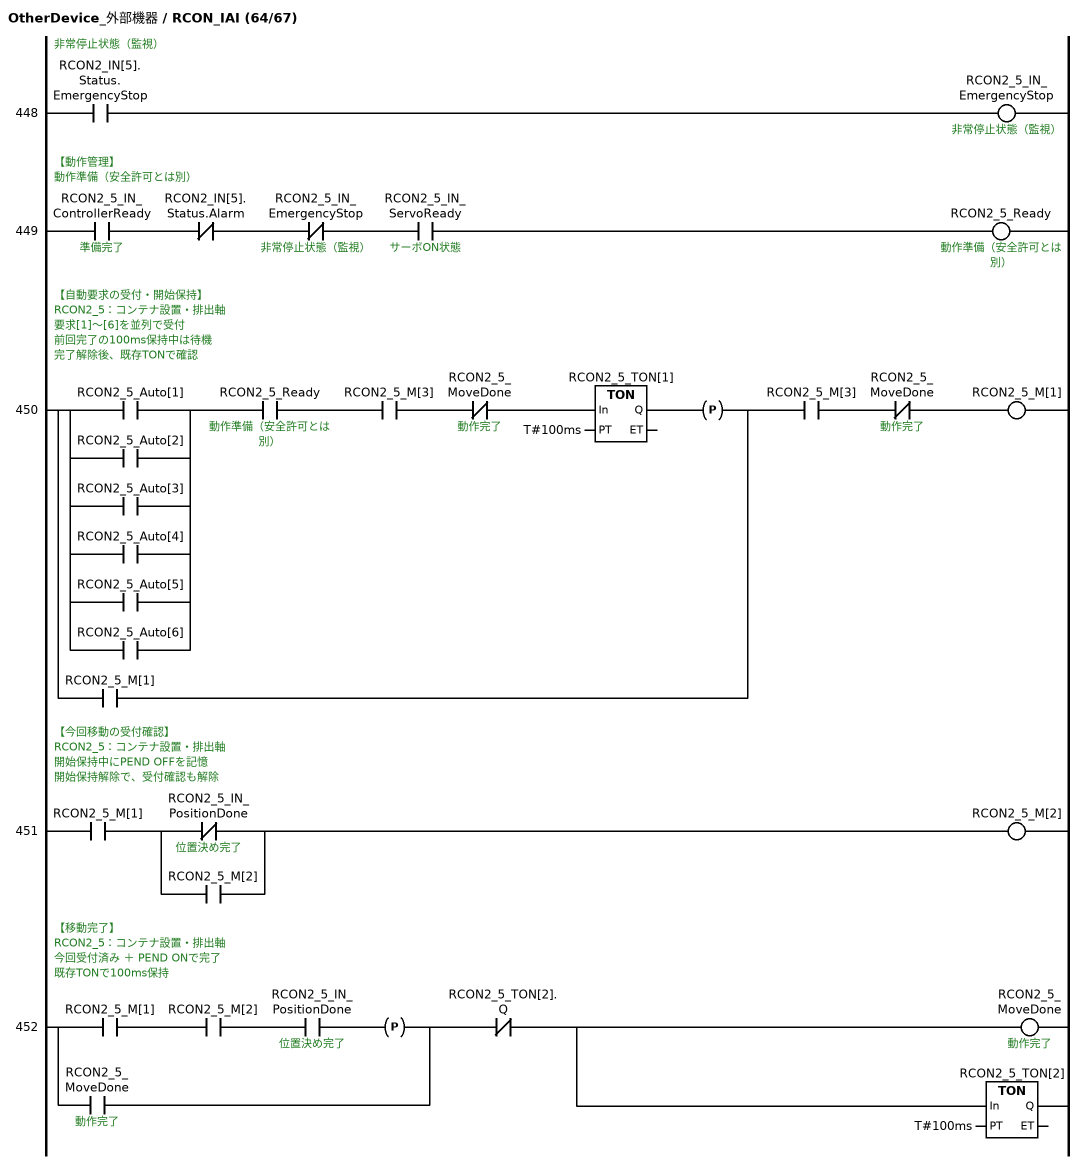
(* Rung 448: 非常停止状態（監視） *)
RCON2_5_IN_EmergencyStop := RCON2_IN[5].Status.EmergencyStop;
(* Rung 449: 【動作管理】 / 動作準備（安全許可とは別） *)
RCON2_5_Ready := RCON2_5_IN_ControllerReady AND NOT RCON2_IN[5].Status.Alarm AND NOT RCON2_5_IN_EmergencyStop AND RCON2_5_IN_ServoReady;
(* Rung 450: 【自動要求の受付・開始保持】 / RCON2_5：コンテナ設置・排出軸 / 要求[1]～[6]を並列で受付 / 前回完了の100ms保持中は待機 / 完了解除後、既存TONで確認 *)
RCON2_5_TON[1](In := (RCON2_5_Auto[1] OR RCON2_5_Auto[2] OR RCON2_5_Auto[3] OR RCON2_5_Auto[4] OR RCON2_5_Auto[5] OR RCON2_5_Auto[6]) AND RCON2_5_Ready AND RCON2_5_M[3] AND NOT RCON2_5_MoveDone, PT := T#100ms);
_e42(CLK := RCON2_5_TON[1].Q);
RCON2_5_M[1] := (_e42.Q OR RCON2_5_M[1]) AND RCON2_5_M[3] AND NOT RCON2_5_MoveDone;
(* Rung 451: 【今回移動の受付確認】 / RCON2_5：コンテナ設置・排出軸 / 開始保持中にPEND OFFを記憶 / 開始保持解除で、受付確認も解除 *)
RCON2_5_M[2] := RCON2_5_M[1] AND (NOT RCON2_5_IN_PositionDone OR RCON2_5_M[2]);
(* Rung 452: 【移動完了】 / RCON2_5：コンテナ設置・排出軸 / 今回受付済み ＋ PEND ONで完了 / 既存TONで100ms保持 *)
_e43(CLK := RCON2_5_M[1] AND RCON2_5_M[2] AND RCON2_5_IN_PositionDone);
_p44 := (_e43.Q OR RCON2_5_MoveDone) AND NOT RCON2_5_TON[2].Q;
RCON2_5_MoveDone := _p44;
RCON2_5_TON[2](In := _p44, PT := T#100ms);

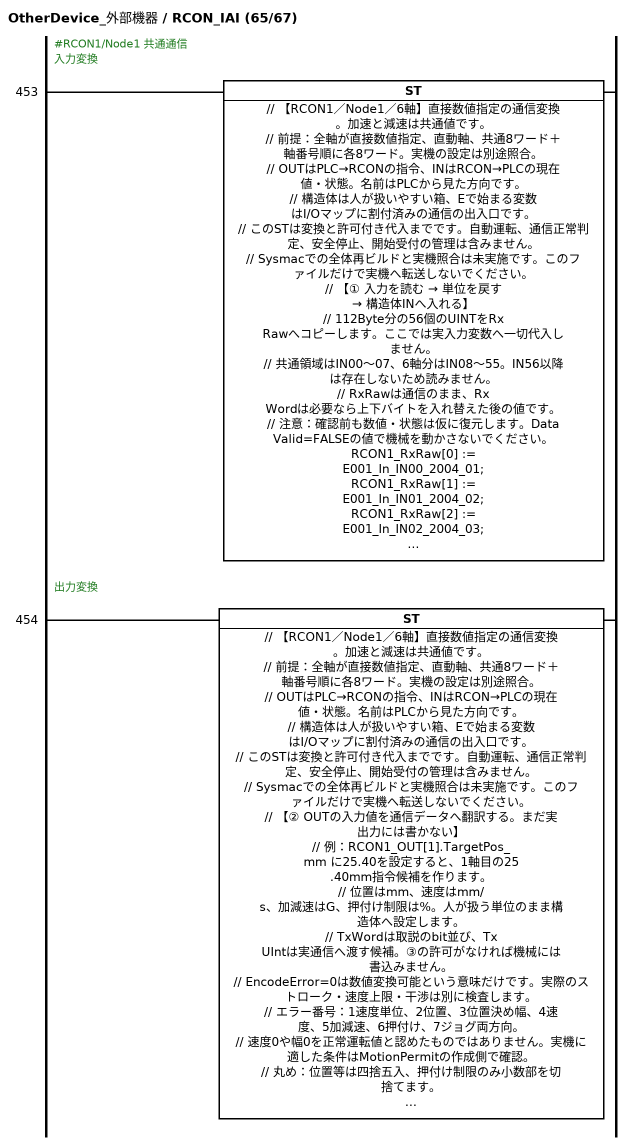
(* Rung 453: #RCON1/Node1 共通通信 / 入力変換 *)
// 【RCON1／Node1／6軸】直接数値指定の通信変換。加速と減速は共通値です。
// 前提：全軸が直接数値指定、直動軸、共通8ワード＋軸番号順に各8ワード。実機の設定は別途照合。
// OUTはPLC→RCONの指令、INはRCON→PLCの現在値・状態。名前はPLCから見た方向です。
// 構造体は人が扱いやすい箱、Eで始まる変数はI/Oマップに割付済みの通信の出入口です。
// このSTは変換と許可付き代入までです。自動運転、通信正常判定、安全停止、開始受付の管理は含みません。
// Sysmacでの全体再ビルドと実機照合は未実施です。このファイルだけで実機へ転送しないでください。
// 【① 入力を読む → 単位を戻す → 構造体INへ入れる】
// 112Byte分の56個のUINTをRxRawへコピーします。ここでは実入力変数へ一切代入しません。
// 共通領域はIN00～07、6軸分はIN08～55。IN56以降は存在しないため読みません。
// RxRawは通信のまま、RxWordは必要なら上下バイトを入れ替えた後の値です。
// 注意：確認前も数値・状態は仮に復元します。DataValid=FALSEの値で機械を動かさないでください。
RCON1_RxRaw[0] := E001_In_IN00_2004_01;
RCON1_RxRaw[1] := E001_In_IN01_2004_02;
RCON1_RxRaw[2] := E001_In_IN02_2004_03;
RCON1_RxRaw[3] := E001_In_IN03_2004_04;
RCON1_RxRaw[4] := E001_In_IN04_2004_05;
RCON1_RxRaw[5] := E001_In_IN05_2004_06;
RCON1_RxRaw[6] := E001_In_IN06_2004_07;
RCON1_RxRaw[7] := E001_In_IN07_2004_08;
RCON1_RxRaw[8] := E001_In_IN08_2004_09;
RCON1_RxRaw[9] := E001_In_IN09_2004_0A;
RCON1_RxRaw[10] := E001_In_IN10_2004_0B;
RCON1_RxRaw[11] := E001_In_IN11_2004_0C;
RCON1_RxRaw[12] := E001_In_IN12_2004_0D;
RCON1_RxRaw[13] := E001_In_IN13_2004_0E;
RCON1_RxRaw[14] := E001_In_IN14_2004_0F;
RCON1_RxRaw[15] := E001_In_IN15_2004_10;
RCON1_RxRaw[16] := E001_In_IN16_2004_11;
RCON1_RxRaw[17] := E001_In_IN17_2004_12;
RCON1_RxRaw[18] := E001_In_IN18_2004_13;
RCON1_RxRaw[19] := E001_In_IN19_2004_14;
RCON1_RxRaw[20] := E001_In_IN20_2004_15;
RCON1_RxRaw[21] := E001_In_IN21_2004_16;
RCON1_RxRaw[22] := E001_In_IN22_2004_17;
RCON1_RxRaw[23] := E001_In_IN23_2004_18;
RCON1_RxRaw[24] := E001_In_IN24_2004_19;
RCON1_RxRaw[25] := E001_In_IN25_2004_1A;
RCON1_RxRaw[26] := E001_In_IN26_2004_1B;
RCON1_RxRaw[27] := E001_In_IN27_2004_1C;
RCON1_RxRaw[28] := E001_In_IN28_2004_1D;
RCON1_RxRaw[29] := E001_In_IN29_2004_1E;
RCON1_RxRaw[30] := E001_In_IN30_2004_1F;
RCON1_RxRaw[31] := E001_In_IN31_2004_20;
RCON1_RxRaw[32] := E001_In_IN32_2004_21;
RCON1_RxRaw[33] := E001_In_IN33_2004_22;
RCON1_RxRaw[34] := E001_In_IN34_2004_23;
RCON1_RxRaw[35] := E001_In_IN35_2004_24;
RCON1_RxRaw[36] := E001_In_IN36_2004_25;
RCON1_RxRaw[37] := E001_In_IN37_2004_26;
RCON1_RxRaw[38] := E001_In_IN38_2004_27;
RCON1_RxRaw[39] := E001_In_IN39_2004_28;
RCON1_RxRaw[40] := E001_In_IN40_2004_29;
RCON1_RxRaw[41] := E001_In_IN41_2004_2A;
RCON1_RxRaw[42] := E001_In_IN42_2004_2B;
RCON1_RxRaw[43] := E001_In_IN43_2004_2C;
RCON1_RxRaw[44] := E001_In_IN44_2004_2D;
RCON1_RxRaw[45] := E001_In_IN45_2004_2E;
RCON1_RxRaw[46] := E001_In_IN46_2004_2F;
RCON1_RxRaw[47] := E001_In_IN47_2004_30;
RCON1_RxRaw[48] := E001_In_IN48_2004_31;
RCON1_RxRaw[49] := E001_In_IN49_2004_32;
RCON1_RxRaw[50] := E001_In_IN50_2004_33;
RCON1_RxRaw[51] := E001_In_IN51_2004_34;
RCON1_RxRaw[52] := E001_In_IN52_2004_35;
RCON1_RxRaw[53] := E001_In_IN53_2004_36;
RCON1_RxRaw[54] := E001_In_IN54_2004_37;
RCON1_RxRaw[55] := E001_In_IN55_2004_38;
// 取説の論理ワードへ正規化。Swapは1ワード内の上下バイト交換です。
// SwapBytesは推測で設定せず、既知の位置とbitで実機照合してください。
FOR ConvWordIndex := INT#0 TO INT#55 DO
    RCON1_RxWord[ConvWordIndex] := UINT_TO_WORD(RCON1_RxRaw[ConvWordIndex]);
    IF RCON1_SwapBytes THEN
        RCON1_RxWord[ConvWordIndex] := Swap(RCON1_RxWord[ConvWordIndex]);
    END_IF;
END_FOR;

ConvUnitOK := (RCON1_SpeedUnit_mm_s = LREAL#1.0) OR
              (RCON1_SpeedUnit_mm_s = LREAL#0.1);

// 【①-2 共通状態】IN00はユニット全体、IN01は各軸のリンク情報です。
// TestABit(ワード, bit番号)は、そのスイッチがONかをBOOLで取り出す命令です。
// 例：IN01のb0は軸No.0→配列[1]、b1は軸No.1→配列[2]。配列番号と実機軸番号は1違います。
// 共通固定領域。ここで使うbit番号は取説の論理bitです（MJ0384 6-24～6-25）。
RCON1_GwRun := TestABit(RCON1_RxWord[0], USINT#15);
RCON1_GwControllerCommLatch := TestABit(RCON1_RxWord[0], USINT#14);
RCON1_GwAxisCommError := TestABit(RCON1_RxWord[0], USINT#13);
RCON1_GwManual := TestABit(RCON1_RxWord[0], USINT#12);
RCON1_GwHeavyAlarm := TestABit(RCON1_RxWord[0], USINT#11);
RCON1_GwLightAlarm := TestABit(RCON1_RxWord[0], USINT#10);
RCON1_GwSystemStop := TestABit(RCON1_RxWord[0], USINT#8);
RCON1_GwAlarmCode := WORD_TO_UINT(RCON1_RxWord[0] AND WORD#16#00FF);
FOR ConvWordIndex := INT#0 TO INT#4 DO
    RCON1_PowerStateRaw[ConvWordIndex] := RCON1_RxWord[ConvWordIndex + INT#2];
END_FOR;

// 【①-3 軸ごとに同じ読取りを繰り返す】
// FORは1～6軸を順番に処理します。ConvBaseはその軸の先頭番号です。
// 計算：8+(軸番号-1)×8。1軸目=8、2軸目=16、3軸目=24。先頭8ワードは共通領域です。
FOR ConvAxisIndex := INT#1 TO INT#6 DO
    ConvBase := INT#8 + (ConvAxisIndex - INT#1) * INT#8;
    RCON1_AxisLinked[ConvAxisIndex] :=
        TestABit(RCON1_RxWord[1], INT_TO_USINT(ConvAxisIndex - INT#1));

// 例：下位2540／上位0なら32bit値2540→25.40mm。
// 上位を16bit左に動かして下位とORで重ねます。SHLが左シフト、ORがビットの合成です。
// 負位置はDWORD_TO_DINTで符号を復元。下位62996／上位65535なら-2540→-25.40mm。
    // 現在位置：下位・上位を結合、符号付き32bitとして解釈、0.01mmをmmへ。
    ConvDWord := SHL(WORD_TO_DWORD(RCON1_RxWord[ConvBase + INT#1]), ULINT#16)
                 OR WORD_TO_DWORD(RCON1_RxWord[ConvBase]);
    RCON1_IN[ConvAxisIndex].ActualPos_mm :=
        DINT_TO_LREAL(DWORD_TO_DINT(ConvDWord)) * LREAL#0.01;

    // 電流：32bitのmA。RCON-PCでは指令電流であり、実測トルクではありません。
    ConvDWord := SHL(WORD_TO_DWORD(RCON1_RxWord[ConvBase + INT#3]), ULINT#16)
                 OR WORD_TO_DWORD(RCON1_RxWord[ConvBase + INT#2]);
    RCON1_IN[ConvAxisIndex].Current_mA := DWORD_TO_DINT(ConvDWord);

    // 現在速度：16bitの負数をINTとして読む。UINTのまま速度にしません。
    IF ConvUnitOK THEN
        RCON1_IN[ConvAxisIndex].ActualSpeed_mm_s :=
            INT_TO_LREAL(WORD_TO_INT(RCON1_RxWord[ConvBase + INT#4])) * RCON1_SpeedUnit_mm_s;
    END_IF;
    // 単位不明のとき速度は前値を保持し、DataValidはFALSEにします。
    // 軸内の+5ワードは予約のため値を使用しません。
    RCON1_IN[ConvAxisIndex].AlarmCode := WORD_TO_UINT(RCON1_RxWord[ConvBase + INT#6]);

// 例：Status.ServoReady=TRUEは「サーボON状態を受信した」という意味。
// OUT側Control.ServoOn=TRUEは「サーボONを要求する」という意味で、指令と結果を区別します。
    // 状態ワード：12個のBOOLへ分解。予約b6,b9～11は使いません。
    RCON1_IN[ConvAxisIndex].Status.PositionDone := TestABit(RCON1_RxWord[ConvBase + INT#7], USINT#0);
    RCON1_IN[ConvAxisIndex].Status.HomeDone := TestABit(RCON1_RxWord[ConvBase + INT#7], USINT#1);
    RCON1_IN[ConvAxisIndex].Status.Moving := TestABit(RCON1_RxWord[ConvBase + INT#7], USINT#2);
    RCON1_IN[ConvAxisIndex].Status.Alarm := TestABit(RCON1_RxWord[ConvBase + INT#7], USINT#3);
    RCON1_IN[ConvAxisIndex].Status.ServoReady := TestABit(RCON1_RxWord[ConvBase + INT#7], USINT#4);
    RCON1_IN[ConvAxisIndex].Status.PushMiss := TestABit(RCON1_RxWord[ConvBase + INT#7], USINT#5);
    RCON1_IN[ConvAxisIndex].Status.OverloadWarning := TestABit(RCON1_RxWord[ConvBase + INT#7], USINT#7);
    RCON1_IN[ConvAxisIndex].Status.CommandDone := TestABit(RCON1_RxWord[ConvBase + INT#7], USINT#8);
    RCON1_IN[ConvAxisIndex].Status.Zone1 := TestABit(RCON1_RxWord[ConvBase + INT#7], USINT#12);
    RCON1_IN[ConvAxisIndex].Status.Zone2 := TestABit(RCON1_RxWord[ConvBase + INT#7], USINT#13);
    RCON1_IN[ConvAxisIndex].Status.ControllerReady := TestABit(RCON1_RxWord[ConvBase + INT#7], USINT#14);
    RCON1_IN[ConvAxisIndex].Status.EmergencyStop := TestABit(RCON1_RxWord[ConvBase + INT#7], USINT#15);

    // DataValidは直接受信bitではなく、今回の内部設計で決めた内部判定です。
    // CommOKはCPUの実通信状態から別途作成。単にTRUE固定にしないでください。
    // DataValidは運転許可や安全保証ではありません。各異常・原点等は別途確認。
    RCON1_IN[ConvAxisIndex].DataValid := RCON1_CommOK AND RCON1_LayoutConfirmed
        AND RCON1_ByteOrderConfirmed AND ConvUnitOK AND RCON1_GwRun
        AND RCON1_AxisLinked[ConvAxisIndex] AND NOT RCON1_GwAxisCommError;
END_FOR;
(* Rung 454: 出力変換 *)
// 【RCON1／Node1／6軸】直接数値指定の通信変換。加速と減速は共通値です。
// 前提：全軸が直接数値指定、直動軸、共通8ワード＋軸番号順に各8ワード。実機の設定は別途照合。
// OUTはPLC→RCONの指令、INはRCON→PLCの現在値・状態。名前はPLCから見た方向です。
// 構造体は人が扱いやすい箱、Eで始まる変数はI/Oマップに割付済みの通信の出入口です。
// このSTは変換と許可付き代入までです。自動運転、通信正常判定、安全停止、開始受付の管理は含みません。
// Sysmacでの全体再ビルドと実機照合は未実施です。このファイルだけで実機へ転送しないでください。
// 【② OUTの入力値を通信データへ翻訳する。まだ実出力には書かない】
// 例：RCON1_OUT[1].TargetPos_mm に25.40を設定すると、1軸目の25.40mm指令候補を作ります。
// 位置はmm、速度はmm/s、加減速はG、押付け制限は%。人が扱う単位のまま構造体へ設定します。
// TxWordは取説のbit並び、TxUIntは実通信へ渡す候補。③の許可がなければ機械には書込みません。
// EncodeError=0は数値変換可能という意味だけです。実際のストローク・速度上限・干渉は別に検査します。
// エラー番号：1速度単位、2位置、3位置決め幅、4速度、5加減速、6押付け、7ジョグ両方向。
// 速度0や幅0を正常運転値と認めたものではありません。実機に適した条件はMotionPermitの作成側で確認。
// 丸め：位置等は四捨五入、押付け制限のみ小数部を切捨てます。

ConvUnitOK := (RCON1_SpeedUnit_mm_s = LREAL#1.0) OR
              (RCON1_SpeedUnit_mm_s = LREAL#0.1);

// 共通制御：MONは論理b15、RTEは論理b13。他のbitは0。
// MONを落とす処理を安全停止として扱わないでください。
RCON1_TxWord[0] := WORD#16#0000;
IF RCON1_GwMON_Request THEN
    RCON1_TxWord[0] := RCON1_TxWord[0] OR WORD#16#8000;
END_IF;
IF RCON1_GwRTE_Request THEN
    RCON1_TxWord[0] := RCON1_TxWord[0] OR WORD#16#2000;
END_IF;

FOR ConvAxisIndex := INT#1 TO INT#6 DO
    ConvBase := INT#8 + (ConvAxisIndex - INT#1) * INT#8;
    RCON1_EncodeError[ConvAxisIndex] := UINT#0;

    // 比較で範囲を確認してから型変換するため、NaN・無限大も変換対象から外れます。
    // 位置・幅9999.99mmはこの案で採用する通信範囲の上限で、実機ストロークではありません。
    IF NOT ConvUnitOK THEN
        RCON1_EncodeError[ConvAxisIndex] := UINT#1;
    ELSIF NOT ((RCON1_OUT[ConvAxisIndex].TargetPos_mm >= LREAL#-9999.99) AND
               (RCON1_OUT[ConvAxisIndex].TargetPos_mm <= LREAL#9999.99)) THEN
        RCON1_EncodeError[ConvAxisIndex] := UINT#2;
    ELSIF NOT ((RCON1_OUT[ConvAxisIndex].PositionBand_mm >= LREAL#0.0) AND
               (RCON1_OUT[ConvAxisIndex].PositionBand_mm <= LREAL#9999.99)) THEN
        RCON1_EncodeError[ConvAxisIndex] := UINT#3;
    ELSIF NOT ((RCON1_OUT[ConvAxisIndex].Speed_mm_s >= LREAL#0.0) AND
               (RCON1_OUT[ConvAxisIndex].Speed_mm_s <= LREAL#65535.0 * RCON1_SpeedUnit_mm_s)) THEN
        RCON1_EncodeError[ConvAxisIndex] := UINT#4;
    ELSIF NOT ((RCON1_OUT[ConvAxisIndex].AccDec_G >= LREAL#0.0) AND
               (RCON1_OUT[ConvAxisIndex].AccDec_G <= LREAL#655.35)) THEN
        RCON1_EncodeError[ConvAxisIndex] := UINT#5;
    ELSIF NOT ((RCON1_OUT[ConvAxisIndex].PushLimit_pct >= LREAL#0.0) AND
               (RCON1_OUT[ConvAxisIndex].PushLimit_pct <= LREAL#200.0)) THEN
        RCON1_EncodeError[ConvAxisIndex] := UINT#6;
    ELSIF RCON1_OUT[ConvAxisIndex].Control.JogMinus AND RCON1_OUT[ConvAxisIndex].Control.JogPlus THEN
        RCON1_EncodeError[ConvAxisIndex] := UINT#7;
    END_IF;

    RCON1_EncodeOK[ConvAxisIndex] := RCON1_EncodeError[ConvAxisIndex] = UINT#0;
    IF RCON1_EncodeOK[ConvAxisIndex] THEN
    // 【数値例】TargetPos_mm=25.40→×100で2540。下位ワード2540、上位ワード0。
// 700.25mm→70025なので下位4489、上位1。65536を超えた分が上位に入ります。
// DINTは符号付きの数、DWORDは同じ32bitの模様。負数の符号を壊さず分割するために使い分けます。
// TRUNCは小数部を捨てます。正数+0.5／負数-0.5を先に行い、四捨五入を明示しています。
    // 目標位置：mmから0.01mmの符号付き整数へ。
        ConvScaled := RCON1_OUT[ConvAxisIndex].TargetPos_mm * LREAL#100.0;
        IF ConvScaled >= LREAL#0.0 THEN
            ConvPos := LINT_TO_DINT(TRUNC(ConvScaled + LREAL#0.5));
        ELSE
            ConvPos := LINT_TO_DINT(TRUNC(ConvScaled - LREAL#0.5));
        END_IF;
        // 負数を含む32bitパターンを保ち、下位・上位の16bitへ分割。
        ConvDWord := DINT_TO_DWORD(ConvPos);
        RCON1_TxWord[ConvBase] := DWORD_TO_WORD(ConvDWord AND DWORD#16#0000FFFF);
        RCON1_TxWord[ConvBase + INT#1] := DWORD_TO_WORD(SHR(ConvDWord, ULINT#16));

        // 位置決め幅：非負の内部整数としてUDINTを選定（メーカーの符号なし保証ではありません）。
        ConvBand := LINT_TO_UDINT(TRUNC(RCON1_OUT[ConvAxisIndex].PositionBand_mm * LREAL#100.0 + LREAL#0.5));
        ConvDWord := UDINT_TO_DWORD(ConvBand);
        RCON1_TxWord[ConvBase + INT#2] := DWORD_TO_WORD(ConvDWord AND DWORD#16#0000FFFF);
        RCON1_TxWord[ConvBase + INT#3] := DWORD_TO_WORD(SHR(ConvDWord, ULINT#16));

// 速度20mm/s：速度単位1.0なら20、0.1なら200を送信します。
// 加減速0.20G：×100して20。加速と減速の両方に同じ値を使います。
// 押付け50%：×255÷100=127.5を切捨てて127。押付けの使用可否・上限は実機仕様で別確認。
        // 速度は1カウント量が1.0か0.1かで値が10倍変わります。
        ConvSpeed := LINT_TO_UINT(TRUNC(RCON1_OUT[ConvAxisIndex].Speed_mm_s / RCON1_SpeedUnit_mm_s + LREAL#0.5));
        ConvAccDec := LINT_TO_UINT(TRUNC(RCON1_OUT[ConvAxisIndex].AccDec_G * LREAL#100.0 + LREAL#0.5));
        ConvPush := LINT_TO_UINT(TRUNC(RCON1_OUT[ConvAxisIndex].PushLimit_pct * LREAL#255.0 / LREAL#100.0));
        RCON1_TxWord[ConvBase + INT#4] := UINT_TO_WORD(ConvSpeed);
        RCON1_TxWord[ConvBase + INT#5] := UINT_TO_WORD(ConvAccDec);
        RCON1_TxWord[ConvBase + INT#6] := UINT_TO_WORD(ConvPush);
    END_IF;
    // 不正値の場合、数値ワードは前値保持。EncodeOK=FALSEで03の書込みを抑止。
    // 前値保持は停止指令ではありません。停止・異常処理は別途設計してください。

    // Controlを論理bitへ詰める。予約b9は必ず0。
    RCON1_TxWord[ConvBase + INT#7] := WORD#16#0000;
// b0 DSTR／Control.Start：TRUEで開始要求。受付応答と10ms以上の保持を確認してOFF。常時ONにしない。
    IF RCON1_OUT[ConvAxisIndex].Control.Start THEN
        RCON1_TxWord[ConvBase + INT#7] := RCON1_TxWord[ConvBase + INT#7] OR WORD#16#0001;
    END_IF;
// b1 HOME／Control.Home：TRUEで原点復帰を指令。原点復帰完了はIN側HomeDoneで確認。
    IF RCON1_OUT[ConvAxisIndex].Control.Home THEN
        RCON1_TxWord[ConvBase + INT#7] := RCON1_TxWord[ConvBase + INT#7] OR WORD#16#0002;
    END_IF;
// b2 STP／Control.Pause：TRUEで一時停止、FALSEで解除。非常停止・安全停止の代用ではない。
    IF RCON1_OUT[ConvAxisIndex].Control.Pause THEN
        RCON1_TxWord[ConvBase + INT#7] := RCON1_TxWord[ConvBase + INT#7] OR WORD#16#0004;
    END_IF;
// b3 RES／Control.Reset：TRUEでアラームリセット要求。コールドスタート級の異常には使用できない。
    IF RCON1_OUT[ConvAxisIndex].Control.Reset THEN
        RCON1_TxWord[ConvBase + INT#7] := RCON1_TxWord[ConvBase + INT#7] OR WORD#16#0008;
    END_IF;
// b4 SON／Control.ServoOn：TRUEでサーボON要求。ON状態はIN側ServoReadyで確認。
    IF RCON1_OUT[ConvAxisIndex].Control.ServoOn THEN
        RCON1_TxWord[ConvBase + INT#7] := RCON1_TxWord[ConvBase + INT#7] OR WORD#16#0010;
    END_IF;
// b5 JISL／Control.InchingSelect：TRUEは一定距離のインチング、FALSEは押している間のジョグ。
    IF RCON1_OUT[ConvAxisIndex].Control.InchingSelect THEN
        RCON1_TxWord[ConvBase + INT#7] := RCON1_TxWord[ConvBase + INT#7] OR WORD#16#0020;
    END_IF;
// b6 JVEL／Control.JogSpeedSelect：FALSEは速度No.26・距離No.48、TRUEは速度No.47または指令速度・距離No.49。
    IF RCON1_OUT[ConvAxisIndex].Control.JogSpeedSelect THEN
        RCON1_TxWord[ConvBase + INT#7] := RCON1_TxWord[ConvBase + INT#7] OR WORD#16#0040;
    END_IF;
// b7 JOG-／Control.JogMinus：TRUEで原点方向へジョグ。反対方向指令との同時ONを防ぐ。
    IF RCON1_OUT[ConvAxisIndex].Control.JogMinus THEN
        RCON1_TxWord[ConvBase + INT#7] := RCON1_TxWord[ConvBase + INT#7] OR WORD#16#0080;
    END_IF;
// b8 JOG+／Control.JogPlus：TRUEで反原点方向へジョグ。反対方向指令との同時ONを防ぐ。
    IF RCON1_OUT[ConvAxisIndex].Control.JogPlus THEN
        RCON1_TxWord[ConvBase + INT#7] := RCON1_TxWord[ConvBase + INT#7] OR WORD#16#0100;
    END_IF;
// b10 GSL0／Control.GainSelect0：GainSelect1と組合せてサーボゲインセット0～3を選ぶ。機械調整用。
    IF RCON1_OUT[ConvAxisIndex].Control.GainSelect0 THEN
        RCON1_TxWord[ConvBase + INT#7] := RCON1_TxWord[ConvBase + INT#7] OR WORD#16#0400;
    END_IF;
// b11 GSL1／Control.GainSelect1：GainSelect0との2bitで選択。速度指令とは別の機能。
    IF RCON1_OUT[ConvAxisIndex].Control.GainSelect1 THEN
        RCON1_TxWord[ConvBase + INT#7] := RCON1_TxWord[ConvBase + INT#7] OR WORD#16#0800;
    END_IF;
// b12 PUSH／Control.PushEnable：TRUEは押付け、FALSEは通常位置決め。押付け条件は別途確認。
    IF RCON1_OUT[ConvAxisIndex].Control.PushEnable THEN
        RCON1_TxWord[ConvBase + INT#7] := RCON1_TxWord[ConvBase + INT#7] OR WORD#16#1000;
    END_IF;
// b13 DIR／Control.PushDirection：CON方式押付け時、TRUEは反原点方向、FALSEは原点方向。
    IF RCON1_OUT[ConvAxisIndex].Control.PushDirection THEN
        RCON1_TxWord[ConvBase + INT#7] := RCON1_TxWord[ConvBase + INT#7] OR WORD#16#2000;
    END_IF;
// b14 INC／Control.RelativeMove：FALSEは絶対座標、TRUEは現在位置からの相対移動量。
    IF RCON1_OUT[ConvAxisIndex].Control.RelativeMove THEN
        RCON1_TxWord[ConvBase + INT#7] := RCON1_TxWord[ConvBase + INT#7] OR WORD#16#4000;
    END_IF;
// b15 BKRL／Control.BrakeRelease：TRUEはブレーキ強制解除。通常FALSE。縦軸では落下等の危険がある。
    IF RCON1_OUT[ConvAxisIndex].Control.BrakeRelease THEN
        RCON1_TxWord[ConvBase + INT#7] := RCON1_TxWord[ConvBase + INT#7] OR WORD#16#8000;
    END_IF;
END_FOR;

// 論理ワードから実際に送るUINTへ。INと同じ1ワード内のバイト交換を適用します。
FOR ConvWordIndex := INT#0 TO INT#55 DO
    ConvWord := RCON1_TxWord[ConvWordIndex];
    IF RCON1_SwapBytes THEN
        ConvWord := Swap(ConvWord);
    END_IF;
    RCON1_TxUInt[ConvWordIndex] := WORD_TO_UINT(ConvWord);
END_FOR;

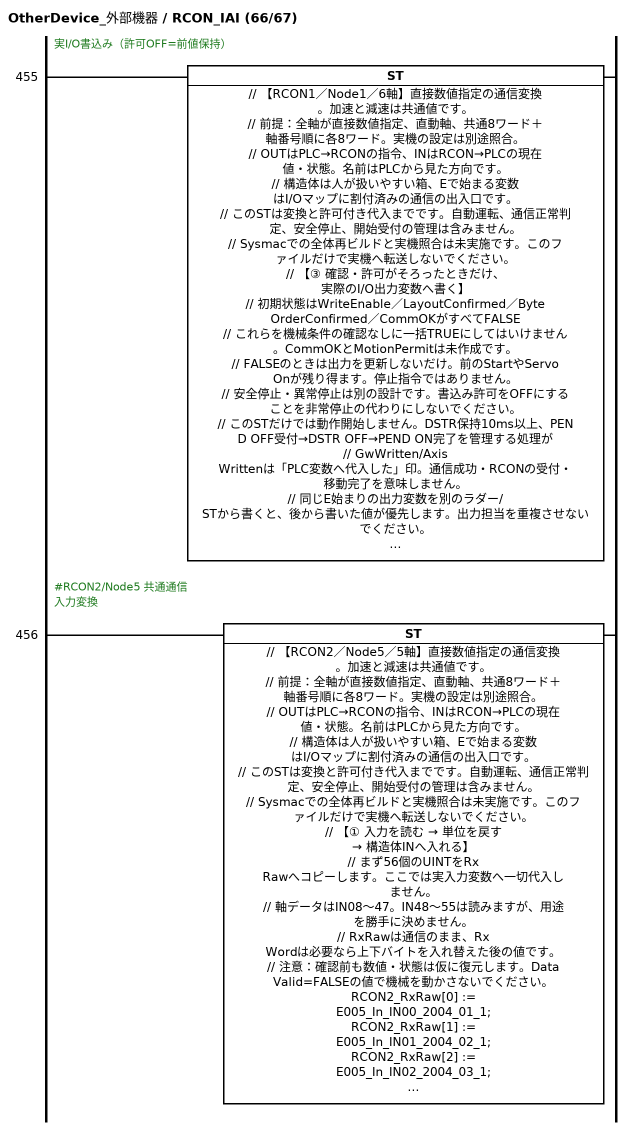
(* Rung 455: 実I/O書込み（許可OFF=前値保持） *)
// 【RCON1／Node1／6軸】直接数値指定の通信変換。加速と減速は共通値です。
// 前提：全軸が直接数値指定、直動軸、共通8ワード＋軸番号順に各8ワード。実機の設定は別途照合。
// OUTはPLC→RCONの指令、INはRCON→PLCの現在値・状態。名前はPLCから見た方向です。
// 構造体は人が扱いやすい箱、Eで始まる変数はI/Oマップに割付済みの通信の出入口です。
// このSTは変換と許可付き代入までです。自動運転、通信正常判定、安全停止、開始受付の管理は含みません。
// Sysmacでの全体再ビルドと実機照合は未実施です。このファイルだけで実機へ転送しないでください。
// 【③ 確認・許可がそろったときだけ、実際のI/O出力変数へ書く】
// 初期状態はWriteEnable／LayoutConfirmed／ByteOrderConfirmed／CommOKがすべてFALSEです。
// これらを機械条件の確認なしに一括TRUEにしてはいけません。CommOKとMotionPermitは未作成です。
// FALSEのときは出力を更新しないだけ。前のStartやServoOnが残り得ます。停止指令ではありません。
// 安全停止・異常停止は別の設計です。書込み許可をOFFにすることを非常停止の代わりにしないでください。
// このSTだけでは動作開始しません。DSTR保持10ms以上、PEND OFF受付→DSTR OFF→PEND ON完了を管理する処理が必要です。
// GwWritten/AxisWrittenは「PLC変数へ代入した」印。通信成功・RCONの受付・移動完了を意味しません。
// 同じE始まりの出力変数を別のラダー/STから書くと、後から書いた値が優先します。出力担当を重複させないでください。

RCON1_GwWritten := FALSE;
FOR ConvAxisIndex := INT#1 TO INT#6 DO
    RCON1_AxisWritten[ConvAxisIndex] := FALSE;
END_FOR;

IF RCON1_WriteEnable AND RCON1_LayoutConfirmed AND RCON1_ByteOrderConfirmed AND RCON1_CommOK THEN
// 共通指令はMON/RTEのみ。最初のRUN応答に必要なため、軸DataValidとは別にGwApplyで許可します。
    IF RCON1_GwApply THEN
        E001_Out_OUT00_2003_01 := RCON1_TxUInt[0];
        RCON1_GwWritten := TRUE;
    END_IF;

// 1軸目＝実機軸No.0。OUT08～OUT15の8ワードをまとめて代入。
// AxisApply=この軸の更新許可、EncodeOK=変換OK、DataValid=入力情報の条件確認、MotionPermit=機械側の運転許可。
// 途中1ワードだけではなく、位置・幅・速度・加減速・押付け・制御を一組として渡します。
    IF RCON1_AxisApply[1] AND RCON1_EncodeOK[1] AND RCON1_IN[1].DataValid
       AND RCON1_MotionPermit[1] THEN
        E001_Out_OUT08_2003_09 := RCON1_TxUInt[8];
        E001_Out_OUT09_2003_0A := RCON1_TxUInt[9];
        E001_Out_OUT10_2003_0B := RCON1_TxUInt[10];
        E001_Out_OUT11_2003_0C := RCON1_TxUInt[11];
        E001_Out_OUT12_2003_0D := RCON1_TxUInt[12];
        E001_Out_OUT13_2003_0E := RCON1_TxUInt[13];
        E001_Out_OUT14_2003_0F := RCON1_TxUInt[14];
        E001_Out_OUT15_2003_10 := RCON1_TxUInt[15];
        RCON1_AxisWritten[1] := TRUE;
    END_IF;

// 2軸目＝実機軸No.1。OUT16～OUT23の8ワードをまとめて代入。
// AxisApply=この軸の更新許可、EncodeOK=変換OK、DataValid=入力情報の条件確認、MotionPermit=機械側の運転許可。
// 途中1ワードだけではなく、位置・幅・速度・加減速・押付け・制御を一組として渡します。
    IF RCON1_AxisApply[2] AND RCON1_EncodeOK[2] AND RCON1_IN[2].DataValid
       AND RCON1_MotionPermit[2] THEN
        E001_Out_OUT16_2003_11 := RCON1_TxUInt[16];
        E001_Out_OUT17_2003_12 := RCON1_TxUInt[17];
        E001_Out_OUT18_2003_13 := RCON1_TxUInt[18];
        E001_Out_OUT19_2003_14 := RCON1_TxUInt[19];
        E001_Out_OUT20_2003_15 := RCON1_TxUInt[20];
        E001_Out_OUT21_2003_16 := RCON1_TxUInt[21];
        E001_Out_OUT22_2003_17 := RCON1_TxUInt[22];
        E001_Out_OUT23_2003_18 := RCON1_TxUInt[23];
        RCON1_AxisWritten[2] := TRUE;
    END_IF;

// 3軸目＝実機軸No.2。OUT24～OUT31の8ワードをまとめて代入。
// AxisApply=この軸の更新許可、EncodeOK=変換OK、DataValid=入力情報の条件確認、MotionPermit=機械側の運転許可。
// 途中1ワードだけではなく、位置・幅・速度・加減速・押付け・制御を一組として渡します。
    IF RCON1_AxisApply[3] AND RCON1_EncodeOK[3] AND RCON1_IN[3].DataValid
       AND RCON1_MotionPermit[3] THEN
        E001_Out_OUT24_2003_19 := RCON1_TxUInt[24];
        E001_Out_OUT25_2003_1A := RCON1_TxUInt[25];
        E001_Out_OUT26_2003_1B := RCON1_TxUInt[26];
        E001_Out_OUT27_2003_1C := RCON1_TxUInt[27];
        E001_Out_OUT28_2003_1D := RCON1_TxUInt[28];
        E001_Out_OUT29_2003_1E := RCON1_TxUInt[29];
        E001_Out_OUT30_2003_1F := RCON1_TxUInt[30];
        E001_Out_OUT31_2003_20 := RCON1_TxUInt[31];
        RCON1_AxisWritten[3] := TRUE;
    END_IF;

// 4軸目＝実機軸No.3。OUT32～OUT39の8ワードをまとめて代入。
// AxisApply=この軸の更新許可、EncodeOK=変換OK、DataValid=入力情報の条件確認、MotionPermit=機械側の運転許可。
// 途中1ワードだけではなく、位置・幅・速度・加減速・押付け・制御を一組として渡します。
    IF RCON1_AxisApply[4] AND RCON1_EncodeOK[4] AND RCON1_IN[4].DataValid
       AND RCON1_MotionPermit[4] THEN
        E001_Out_OUT32_2003_21 := RCON1_TxUInt[32];
        E001_Out_OUT33_2003_22 := RCON1_TxUInt[33];
        E001_Out_OUT34_2003_23 := RCON1_TxUInt[34];
        E001_Out_OUT35_2003_24 := RCON1_TxUInt[35];
        E001_Out_OUT36_2003_25 := RCON1_TxUInt[36];
        E001_Out_OUT37_2003_26 := RCON1_TxUInt[37];
        E001_Out_OUT38_2003_27 := RCON1_TxUInt[38];
        E001_Out_OUT39_2003_28 := RCON1_TxUInt[39];
        RCON1_AxisWritten[4] := TRUE;
    END_IF;

// 5軸目＝実機軸No.4。OUT40～OUT47の8ワードをまとめて代入。
// AxisApply=この軸の更新許可、EncodeOK=変換OK、DataValid=入力情報の条件確認、MotionPermit=機械側の運転許可。
// 途中1ワードだけではなく、位置・幅・速度・加減速・押付け・制御を一組として渡します。
    IF RCON1_AxisApply[5] AND RCON1_EncodeOK[5] AND RCON1_IN[5].DataValid
       AND RCON1_MotionPermit[5] THEN
        E001_Out_OUT40_2003_29 := RCON1_TxUInt[40];
        E001_Out_OUT41_2003_2A := RCON1_TxUInt[41];
        E001_Out_OUT42_2003_2B := RCON1_TxUInt[42];
        E001_Out_OUT43_2003_2C := RCON1_TxUInt[43];
        E001_Out_OUT44_2003_2D := RCON1_TxUInt[44];
        E001_Out_OUT45_2003_2E := RCON1_TxUInt[45];
        E001_Out_OUT46_2003_2F := RCON1_TxUInt[46];
        E001_Out_OUT47_2003_30 := RCON1_TxUInt[47];
        RCON1_AxisWritten[5] := TRUE;
    END_IF;

// 6軸目＝実機軸No.5。OUT48～OUT55の8ワードをまとめて代入。
// AxisApply=この軸の更新許可、EncodeOK=変換OK、DataValid=入力情報の条件確認、MotionPermit=機械側の運転許可。
// 途中1ワードだけではなく、位置・幅・速度・加減速・押付け・制御を一組として渡します。
    IF RCON1_AxisApply[6] AND RCON1_EncodeOK[6] AND RCON1_IN[6].DataValid
       AND RCON1_MotionPermit[6] THEN
        E001_Out_OUT48_2003_31 := RCON1_TxUInt[48];
        E001_Out_OUT49_2003_32 := RCON1_TxUInt[49];
        E001_Out_OUT50_2003_33 := RCON1_TxUInt[50];
        E001_Out_OUT51_2003_34 := RCON1_TxUInt[51];
        E001_Out_OUT52_2003_35 := RCON1_TxUInt[52];
        E001_Out_OUT53_2003_36 := RCON1_TxUInt[53];
        E001_Out_OUT54_2003_37 := RCON1_TxUInt[54];
        E001_Out_OUT55_2003_38 := RCON1_TxUInt[55];
        RCON1_AxisWritten[6] := TRUE;
    END_IF;
END_IF;
// OUT01～07は予約領域のため書き換えません。OUT56以降は112Byte設定に存在しません。
// 現在の実機設定・別処理の用途が未確認なので、余剰領域を勝手にゼロクリアしません。
(* Rung 456: #RCON2/Node5 共通通信 / 入力変換 *)
// 【RCON2／Node5／5軸】直接数値指定の通信変換。加速と減速は共通値です。
// 前提：全軸が直接数値指定、直動軸、共通8ワード＋軸番号順に各8ワード。実機の設定は別途照合。
// OUTはPLC→RCONの指令、INはRCON→PLCの現在値・状態。名前はPLCから見た方向です。
// 構造体は人が扱いやすい箱、Eで始まる変数はI/Oマップに割付済みの通信の出入口です。
// このSTは変換と許可付き代入までです。自動運転、通信正常判定、安全停止、開始受付の管理は含みません。
// Sysmacでの全体再ビルドと実機照合は未実施です。このファイルだけで実機へ転送しないでください。
// 【① 入力を読む → 単位を戻す → 構造体INへ入れる】
// まず56個のUINTをRxRawへコピーします。ここでは実入力変数へ一切代入しません。
// 軸データはIN08～47。IN48～55は読みますが、用途を勝手に決めません。
// RxRawは通信のまま、RxWordは必要なら上下バイトを入れ替えた後の値です。
// 注意：確認前も数値・状態は仮に復元します。DataValid=FALSEの値で機械を動かさないでください。
RCON2_RxRaw[0] := E005_In_IN00_2004_01_1;
RCON2_RxRaw[1] := E005_In_IN01_2004_02_1;
RCON2_RxRaw[2] := E005_In_IN02_2004_03_1;
RCON2_RxRaw[3] := E005_In_IN03_2004_04_1;
RCON2_RxRaw[4] := E005_In_IN04_2004_05_1;
RCON2_RxRaw[5] := E005_In_IN05_2004_06_1;
RCON2_RxRaw[6] := E005_In_IN06_2004_07_1;
RCON2_RxRaw[7] := E005_In_IN07_2004_08_1;
RCON2_RxRaw[8] := E005_In_IN08_2004_09_1;
RCON2_RxRaw[9] := E005_In_IN09_2004_0A_1;
RCON2_RxRaw[10] := E005_In_IN10_2004_0B_1;
RCON2_RxRaw[11] := E005_In_IN11_2004_0C_1;
RCON2_RxRaw[12] := E005_In_IN12_2004_0D_1;
RCON2_RxRaw[13] := E005_In_IN13_2004_0E_1;
RCON2_RxRaw[14] := E005_In_IN14_2004_0F_1;
RCON2_RxRaw[15] := E005_In_IN15_2004_10_1;
RCON2_RxRaw[16] := E005_In_IN16_2004_11_1;
RCON2_RxRaw[17] := E005_In_IN17_2004_12_1;
RCON2_RxRaw[18] := E005_In_IN18_2004_13_1;
RCON2_RxRaw[19] := E005_In_IN19_2004_14_1;
RCON2_RxRaw[20] := E005_In_IN20_2004_15_1;
RCON2_RxRaw[21] := E005_In_IN21_2004_16_1;
RCON2_RxRaw[22] := E005_In_IN22_2004_17_1;
RCON2_RxRaw[23] := E005_In_IN23_2004_18_1;
RCON2_RxRaw[24] := E005_In_IN24_2004_19_1;
RCON2_RxRaw[25] := E005_In_IN25_2004_1A_1;
RCON2_RxRaw[26] := E005_In_IN26_2004_1B_1;
RCON2_RxRaw[27] := E005_In_IN27_2004_1C_1;
RCON2_RxRaw[28] := E005_In_IN28_2004_1D_1;
RCON2_RxRaw[29] := E005_In_IN29_2004_1E_1;
RCON2_RxRaw[30] := E005_In_IN30_2004_1F_1;
RCON2_RxRaw[31] := E005_In_IN31_2004_20_1;
RCON2_RxRaw[32] := E005_In_IN32_2004_21_1;
RCON2_RxRaw[33] := E005_In_IN33_2004_22_1;
RCON2_RxRaw[34] := E005_In_IN34_2004_23_1;
RCON2_RxRaw[35] := E005_In_IN35_2004_24_1;
RCON2_RxRaw[36] := E005_In_IN36_2004_25_1;
RCON2_RxRaw[37] := E005_In_IN37_2004_26_1;
RCON2_RxRaw[38] := E005_In_IN38_2004_27_1;
RCON2_RxRaw[39] := E005_In_IN39_2004_28_1;
RCON2_RxRaw[40] := E005_In_IN40_2004_29_1;
RCON2_RxRaw[41] := E005_In_IN41_2004_2A_1;
RCON2_RxRaw[42] := E005_In_IN42_2004_2B_1;
RCON2_RxRaw[43] := E005_In_IN43_2004_2C_1;
RCON2_RxRaw[44] := E005_In_IN44_2004_2D_1;
RCON2_RxRaw[45] := E005_In_IN45_2004_2E_1;
RCON2_RxRaw[46] := E005_In_IN46_2004_2F_1;
RCON2_RxRaw[47] := E005_In_IN47_2004_30_1;
RCON2_RxRaw[48] := E005_In_IN48_2004_31_1;
RCON2_RxRaw[49] := E005_In_IN49_2004_32_1;
RCON2_RxRaw[50] := E005_In_IN50_2004_33_1;
RCON2_RxRaw[51] := E005_In_IN51_2004_34_1;
RCON2_RxRaw[52] := E005_In_IN52_2004_35_1;
RCON2_RxRaw[53] := E005_In_IN53_2004_36_1;
RCON2_RxRaw[54] := E005_In_IN54_2004_37_1;
RCON2_RxRaw[55] := E005_In_IN55_2004_38_1;

// 取説の論理ワードへ正規化。Swapは1ワード内の上下バイト交換です。
// SwapBytesは推測で設定せず、既知の位置とbitで実機照合してください。
FOR ConvWordIndex := INT#0 TO INT#55 DO
    RCON2_RxWord[ConvWordIndex] := UINT_TO_WORD(RCON2_RxRaw[ConvWordIndex]);
    IF RCON2_SwapBytes THEN
        RCON2_RxWord[ConvWordIndex] := Swap(RCON2_RxWord[ConvWordIndex]);
    END_IF;
END_FOR;

ConvUnitOK := (RCON2_SpeedUnit_mm_s = LREAL#1.0) OR
              (RCON2_SpeedUnit_mm_s = LREAL#0.1);

// 【①-2 共通状態】IN00はユニット全体、IN01は各軸のリンク情報です。
// TestABit(ワード, bit番号)は、そのスイッチがONかをBOOLで取り出す命令です。
// 例：IN01のb0は軸No.0→配列[1]、b1は軸No.1→配列[2]。配列番号と実機軸番号は1違います。
// 共通固定領域。ここで使うbit番号は取説の論理bitです（MJ0384 6-24～6-25）。
RCON2_GwRun := TestABit(RCON2_RxWord[0], USINT#15);
RCON2_GwControllerCommLatch := TestABit(RCON2_RxWord[0], USINT#14);
RCON2_GwAxisCommError := TestABit(RCON2_RxWord[0], USINT#13);
RCON2_GwManual := TestABit(RCON2_RxWord[0], USINT#12);
RCON2_GwHeavyAlarm := TestABit(RCON2_RxWord[0], USINT#11);
RCON2_GwLightAlarm := TestABit(RCON2_RxWord[0], USINT#10);
RCON2_GwSystemStop := TestABit(RCON2_RxWord[0], USINT#8);
RCON2_GwAlarmCode := WORD_TO_UINT(RCON2_RxWord[0] AND WORD#16#00FF);
FOR ConvWordIndex := INT#0 TO INT#4 DO
    RCON2_PowerStateRaw[ConvWordIndex] := RCON2_RxWord[ConvWordIndex + INT#2];
END_FOR;

// 【①-3 軸ごとに同じ読取りを繰り返す】
// FORは1～5軸を順番に処理します。ConvBaseはその軸の先頭番号です。
// 計算：8+(軸番号-1)×8。1軸目=8、2軸目=16、3軸目=24。先頭8ワードは共通領域です。
FOR ConvAxisIndex := INT#1 TO INT#5 DO
    ConvBase := INT#8 + (ConvAxisIndex - INT#1) * INT#8;
    RCON2_AxisLinked[ConvAxisIndex] :=
        TestABit(RCON2_RxWord[1], INT_TO_USINT(ConvAxisIndex - INT#1));

// 例：下位2540／上位0なら32bit値2540→25.40mm。
// 上位を16bit左に動かして下位とORで重ねます。SHLが左シフト、ORがビットの合成です。
// 負位置はDWORD_TO_DINTで符号を復元。下位62996／上位65535なら-2540→-25.40mm。
    // 現在位置：下位・上位を結合、符号付き32bitとして解釈、0.01mmをmmへ。
    ConvDWord := SHL(WORD_TO_DWORD(RCON2_RxWord[ConvBase + INT#1]), ULINT#16)
                 OR WORD_TO_DWORD(RCON2_RxWord[ConvBase]);
    RCON2_IN[ConvAxisIndex].ActualPos_mm :=
        DINT_TO_LREAL(DWORD_TO_DINT(ConvDWord)) * LREAL#0.01;

    // 電流：32bitのmA。RCON-PCでは指令電流であり、実測トルクではありません。
    ConvDWord := SHL(WORD_TO_DWORD(RCON2_RxWord[ConvBase + INT#3]), ULINT#16)
                 OR WORD_TO_DWORD(RCON2_RxWord[ConvBase + INT#2]);
    RCON2_IN[ConvAxisIndex].Current_mA := DWORD_TO_DINT(ConvDWord);

    // 現在速度：16bitの負数をINTとして読む。UINTのまま速度にしません。
    IF ConvUnitOK THEN
        RCON2_IN[ConvAxisIndex].ActualSpeed_mm_s :=
            INT_TO_LREAL(WORD_TO_INT(RCON2_RxWord[ConvBase + INT#4])) * RCON2_SpeedUnit_mm_s;
    END_IF;
    // 単位不明のとき速度は前値を保持し、DataValidはFALSEにします。
    // 軸内の+5ワードは予約のため値を使用しません。
    RCON2_IN[ConvAxisIndex].AlarmCode := WORD_TO_UINT(RCON2_RxWord[ConvBase + INT#6]);

// 例：Status.ServoReady=TRUEは「サーボON状態を受信した」という意味。
// OUT側Control.ServoOn=TRUEは「サーボONを要求する」という意味で、指令と結果を区別します。
    // 状態ワード：12個のBOOLへ分解。予約b6,b9～11は使いません。
    RCON2_IN[ConvAxisIndex].Status.PositionDone := TestABit(RCON2_RxWord[ConvBase + INT#7], USINT#0);
    RCON2_IN[ConvAxisIndex].Status.HomeDone := TestABit(RCON2_RxWord[ConvBase + INT#7], USINT#1);
    RCON2_IN[ConvAxisIndex].Status.Moving := TestABit(RCON2_RxWord[ConvBase + INT#7], USINT#2);
    RCON2_IN[ConvAxisIndex].Status.Alarm := TestABit(RCON2_RxWord[ConvBase + INT#7], USINT#3);
    RCON2_IN[ConvAxisIndex].Status.ServoReady := TestABit(RCON2_RxWord[ConvBase + INT#7], USINT#4);
    RCON2_IN[ConvAxisIndex].Status.PushMiss := TestABit(RCON2_RxWord[ConvBase + INT#7], USINT#5);
    RCON2_IN[ConvAxisIndex].Status.OverloadWarning := TestABit(RCON2_RxWord[ConvBase + INT#7], USINT#7);
    RCON2_IN[ConvAxisIndex].Status.CommandDone := TestABit(RCON2_RxWord[ConvBase + INT#7], USINT#8);
    RCON2_IN[ConvAxisIndex].Status.Zone1 := TestABit(RCON2_RxWord[ConvBase + INT#7], USINT#12);
    RCON2_IN[ConvAxisIndex].Status.Zone2 := TestABit(RCON2_RxWord[ConvBase + INT#7], USINT#13);
    RCON2_IN[ConvAxisIndex].Status.ControllerReady := TestABit(RCON2_RxWord[ConvBase + INT#7], USINT#14);
    RCON2_IN[ConvAxisIndex].Status.EmergencyStop := TestABit(RCON2_RxWord[ConvBase + INT#7], USINT#15);

    // DataValidは直接受信bitではなく、今回の内部設計で決めた内部判定です。
    // CommOKはCPUの実通信状態から別途作成。単にTRUE固定にしないでください。
    // DataValidは運転許可や安全保証ではありません。各異常・原点等は別途確認。
    RCON2_IN[ConvAxisIndex].DataValid := RCON2_CommOK AND RCON2_LayoutConfirmed
        AND RCON2_ByteOrderConfirmed AND ConvUnitOK AND RCON2_GwRun
        AND RCON2_AxisLinked[ConvAxisIndex] AND NOT RCON2_GwAxisCommError;
END_FOR;

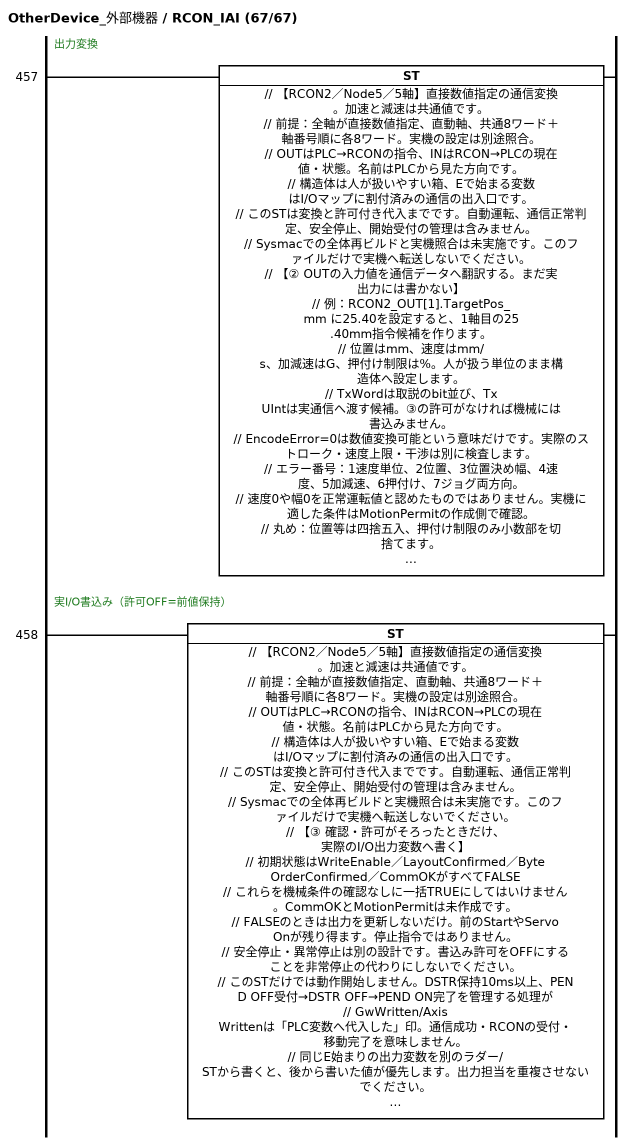
(* Rung 457: 出力変換 *)
// 【RCON2／Node5／5軸】直接数値指定の通信変換。加速と減速は共通値です。
// 前提：全軸が直接数値指定、直動軸、共通8ワード＋軸番号順に各8ワード。実機の設定は別途照合。
// OUTはPLC→RCONの指令、INはRCON→PLCの現在値・状態。名前はPLCから見た方向です。
// 構造体は人が扱いやすい箱、Eで始まる変数はI/Oマップに割付済みの通信の出入口です。
// このSTは変換と許可付き代入までです。自動運転、通信正常判定、安全停止、開始受付の管理は含みません。
// Sysmacでの全体再ビルドと実機照合は未実施です。このファイルだけで実機へ転送しないでください。
// 【② OUTの入力値を通信データへ翻訳する。まだ実出力には書かない】
// 例：RCON2_OUT[1].TargetPos_mm に25.40を設定すると、1軸目の25.40mm指令候補を作ります。
// 位置はmm、速度はmm/s、加減速はG、押付け制限は%。人が扱う単位のまま構造体へ設定します。
// TxWordは取説のbit並び、TxUIntは実通信へ渡す候補。③の許可がなければ機械には書込みません。
// EncodeError=0は数値変換可能という意味だけです。実際のストローク・速度上限・干渉は別に検査します。
// エラー番号：1速度単位、2位置、3位置決め幅、4速度、5加減速、6押付け、7ジョグ両方向。
// 速度0や幅0を正常運転値と認めたものではありません。実機に適した条件はMotionPermitの作成側で確認。
// 丸め：位置等は四捨五入、押付け制限のみ小数部を切捨てます。

ConvUnitOK := (RCON2_SpeedUnit_mm_s = LREAL#1.0) OR
              (RCON2_SpeedUnit_mm_s = LREAL#0.1);

// 共通制御：MONは論理b15、RTEは論理b13。他のbitは0。
// MONを落とす処理を安全停止として扱わないでください。
RCON2_TxWord[0] := WORD#16#0000;
IF RCON2_GwMON_Request THEN
    RCON2_TxWord[0] := RCON2_TxWord[0] OR WORD#16#8000;
END_IF;
IF RCON2_GwRTE_Request THEN
    RCON2_TxWord[0] := RCON2_TxWord[0] OR WORD#16#2000;
END_IF;

FOR ConvAxisIndex := INT#1 TO INT#5 DO
    ConvBase := INT#8 + (ConvAxisIndex - INT#1) * INT#8;
    RCON2_EncodeError[ConvAxisIndex] := UINT#0;

    // 比較で範囲を確認してから型変換するため、NaN・無限大も変換対象から外れます。
    // 位置・幅9999.99mmはこの案で採用する通信範囲の上限で、実機ストロークではありません。
    IF NOT ConvUnitOK THEN
        RCON2_EncodeError[ConvAxisIndex] := UINT#1;
    ELSIF NOT ((RCON2_OUT[ConvAxisIndex].TargetPos_mm >= LREAL#-9999.99) AND
               (RCON2_OUT[ConvAxisIndex].TargetPos_mm <= LREAL#9999.99)) THEN
        RCON2_EncodeError[ConvAxisIndex] := UINT#2;
    ELSIF NOT ((RCON2_OUT[ConvAxisIndex].PositionBand_mm >= LREAL#0.0) AND
               (RCON2_OUT[ConvAxisIndex].PositionBand_mm <= LREAL#9999.99)) THEN
        RCON2_EncodeError[ConvAxisIndex] := UINT#3;
    ELSIF NOT ((RCON2_OUT[ConvAxisIndex].Speed_mm_s >= LREAL#0.0) AND
               (RCON2_OUT[ConvAxisIndex].Speed_mm_s <= LREAL#65535.0 * RCON2_SpeedUnit_mm_s)) THEN
        RCON2_EncodeError[ConvAxisIndex] := UINT#4;
    ELSIF NOT ((RCON2_OUT[ConvAxisIndex].AccDec_G >= LREAL#0.0) AND
               (RCON2_OUT[ConvAxisIndex].AccDec_G <= LREAL#655.35)) THEN
        RCON2_EncodeError[ConvAxisIndex] := UINT#5;
    ELSIF NOT ((RCON2_OUT[ConvAxisIndex].PushLimit_pct >= LREAL#0.0) AND
               (RCON2_OUT[ConvAxisIndex].PushLimit_pct <= LREAL#200.0)) THEN
        RCON2_EncodeError[ConvAxisIndex] := UINT#6;
    ELSIF RCON2_OUT[ConvAxisIndex].Control.JogMinus AND RCON2_OUT[ConvAxisIndex].Control.JogPlus THEN
        RCON2_EncodeError[ConvAxisIndex] := UINT#7;
    END_IF;

    RCON2_EncodeOK[ConvAxisIndex] := RCON2_EncodeError[ConvAxisIndex] = UINT#0;
    IF RCON2_EncodeOK[ConvAxisIndex] THEN
    // 【数値例】TargetPos_mm=25.40→×100で2540。下位ワード2540、上位ワード0。
// 700.25mm→70025なので下位4489、上位1。65536を超えた分が上位に入ります。
// DINTは符号付きの数、DWORDは同じ32bitの模様。負数の符号を壊さず分割するために使い分けます。
// TRUNCは小数部を捨てます。正数+0.5／負数-0.5を先に行い、四捨五入を明示しています。
    // 目標位置：mmから0.01mmの符号付き整数へ。
        ConvScaled := RCON2_OUT[ConvAxisIndex].TargetPos_mm * LREAL#100.0;
        IF ConvScaled >= LREAL#0.0 THEN
            ConvPos := LINT_TO_DINT(TRUNC(ConvScaled + LREAL#0.5));
        ELSE
            ConvPos := LINT_TO_DINT(TRUNC(ConvScaled - LREAL#0.5));
        END_IF;
        // 負数を含む32bitパターンを保ち、下位・上位の16bitへ分割。
        ConvDWord := DINT_TO_DWORD(ConvPos);
        RCON2_TxWord[ConvBase] := DWORD_TO_WORD(ConvDWord AND DWORD#16#0000FFFF);
        RCON2_TxWord[ConvBase + INT#1] := DWORD_TO_WORD(SHR(ConvDWord, ULINT#16));

        // 位置決め幅：非負の内部整数としてUDINTを選定（メーカーの符号なし保証ではありません）。
        ConvBand := LINT_TO_UDINT(TRUNC(RCON2_OUT[ConvAxisIndex].PositionBand_mm * LREAL#100.0 + LREAL#0.5));
        ConvDWord := UDINT_TO_DWORD(ConvBand);
        RCON2_TxWord[ConvBase + INT#2] := DWORD_TO_WORD(ConvDWord AND DWORD#16#0000FFFF);
        RCON2_TxWord[ConvBase + INT#3] := DWORD_TO_WORD(SHR(ConvDWord, ULINT#16));

// 速度20mm/s：速度単位1.0なら20、0.1なら200を送信します。
// 加減速0.20G：×100して20。加速と減速の両方に同じ値を使います。
// 押付け50%：×255÷100=127.5を切捨てて127。押付けの使用可否・上限は実機仕様で別確認。
        // 速度は1カウント量が1.0か0.1かで値が10倍変わります。
        ConvSpeed := LINT_TO_UINT(TRUNC(RCON2_OUT[ConvAxisIndex].Speed_mm_s / RCON2_SpeedUnit_mm_s + LREAL#0.5));
        ConvAccDec := LINT_TO_UINT(TRUNC(RCON2_OUT[ConvAxisIndex].AccDec_G * LREAL#100.0 + LREAL#0.5));
        ConvPush := LINT_TO_UINT(TRUNC(RCON2_OUT[ConvAxisIndex].PushLimit_pct * LREAL#255.0 / LREAL#100.0));
        RCON2_TxWord[ConvBase + INT#4] := UINT_TO_WORD(ConvSpeed);
        RCON2_TxWord[ConvBase + INT#5] := UINT_TO_WORD(ConvAccDec);
        RCON2_TxWord[ConvBase + INT#6] := UINT_TO_WORD(ConvPush);
    END_IF;
    // 不正値の場合、数値ワードは前値保持。EncodeOK=FALSEで03の書込みを抑止。
    // 前値保持は停止指令ではありません。停止・異常処理は別途設計してください。

    // Controlを論理bitへ詰める。予約b9は必ず0。
    RCON2_TxWord[ConvBase + INT#7] := WORD#16#0000;
// b0 DSTR／Control.Start：TRUEで開始要求。受付応答と10ms以上の保持を確認してOFF。常時ONにしない。
    IF RCON2_OUT[ConvAxisIndex].Control.Start THEN
        RCON2_TxWord[ConvBase + INT#7] := RCON2_TxWord[ConvBase + INT#7] OR WORD#16#0001;
    END_IF;
// b1 HOME／Control.Home：TRUEで原点復帰を指令。原点復帰完了はIN側HomeDoneで確認。
    IF RCON2_OUT[ConvAxisIndex].Control.Home THEN
        RCON2_TxWord[ConvBase + INT#7] := RCON2_TxWord[ConvBase + INT#7] OR WORD#16#0002;
    END_IF;
// b2 STP／Control.Pause：TRUEで一時停止、FALSEで解除。非常停止・安全停止の代用ではない。
    IF RCON2_OUT[ConvAxisIndex].Control.Pause THEN
        RCON2_TxWord[ConvBase + INT#7] := RCON2_TxWord[ConvBase + INT#7] OR WORD#16#0004;
    END_IF;
// b3 RES／Control.Reset：TRUEでアラームリセット要求。コールドスタート級の異常には使用できない。
    IF RCON2_OUT[ConvAxisIndex].Control.Reset THEN
        RCON2_TxWord[ConvBase + INT#7] := RCON2_TxWord[ConvBase + INT#7] OR WORD#16#0008;
    END_IF;
// b4 SON／Control.ServoOn：TRUEでサーボON要求。ON状態はIN側ServoReadyで確認。
    IF RCON2_OUT[ConvAxisIndex].Control.ServoOn THEN
        RCON2_TxWord[ConvBase + INT#7] := RCON2_TxWord[ConvBase + INT#7] OR WORD#16#0010;
    END_IF;
// b5 JISL／Control.InchingSelect：TRUEは一定距離のインチング、FALSEは押している間のジョグ。
    IF RCON2_OUT[ConvAxisIndex].Control.InchingSelect THEN
        RCON2_TxWord[ConvBase + INT#7] := RCON2_TxWord[ConvBase + INT#7] OR WORD#16#0020;
    END_IF;
// b6 JVEL／Control.JogSpeedSelect：FALSEは速度No.26・距離No.48、TRUEは速度No.47または指令速度・距離No.49。
    IF RCON2_OUT[ConvAxisIndex].Control.JogSpeedSelect THEN
        RCON2_TxWord[ConvBase + INT#7] := RCON2_TxWord[ConvBase + INT#7] OR WORD#16#0040;
    END_IF;
// b7 JOG-／Control.JogMinus：TRUEで原点方向へジョグ。反対方向指令との同時ONを防ぐ。
    IF RCON2_OUT[ConvAxisIndex].Control.JogMinus THEN
        RCON2_TxWord[ConvBase + INT#7] := RCON2_TxWord[ConvBase + INT#7] OR WORD#16#0080;
    END_IF;
// b8 JOG+／Control.JogPlus：TRUEで反原点方向へジョグ。反対方向指令との同時ONを防ぐ。
    IF RCON2_OUT[ConvAxisIndex].Control.JogPlus THEN
        RCON2_TxWord[ConvBase + INT#7] := RCON2_TxWord[ConvBase + INT#7] OR WORD#16#0100;
    END_IF;
// b10 GSL0／Control.GainSelect0：GainSelect1と組合せてサーボゲインセット0～3を選ぶ。機械調整用。
    IF RCON2_OUT[ConvAxisIndex].Control.GainSelect0 THEN
        RCON2_TxWord[ConvBase + INT#7] := RCON2_TxWord[ConvBase + INT#7] OR WORD#16#0400;
    END_IF;
// b11 GSL1／Control.GainSelect1：GainSelect0との2bitで選択。速度指令とは別の機能。
    IF RCON2_OUT[ConvAxisIndex].Control.GainSelect1 THEN
        RCON2_TxWord[ConvBase + INT#7] := RCON2_TxWord[ConvBase + INT#7] OR WORD#16#0800;
    END_IF;
// b12 PUSH／Control.PushEnable：TRUEは押付け、FALSEは通常位置決め。押付け条件は別途確認。
    IF RCON2_OUT[ConvAxisIndex].Control.PushEnable THEN
        RCON2_TxWord[ConvBase + INT#7] := RCON2_TxWord[ConvBase + INT#7] OR WORD#16#1000;
    END_IF;
// b13 DIR／Control.PushDirection：CON方式押付け時、TRUEは反原点方向、FALSEは原点方向。
    IF RCON2_OUT[ConvAxisIndex].Control.PushDirection THEN
        RCON2_TxWord[ConvBase + INT#7] := RCON2_TxWord[ConvBase + INT#7] OR WORD#16#2000;
    END_IF;
// b14 INC／Control.RelativeMove：FALSEは絶対座標、TRUEは現在位置からの相対移動量。
    IF RCON2_OUT[ConvAxisIndex].Control.RelativeMove THEN
        RCON2_TxWord[ConvBase + INT#7] := RCON2_TxWord[ConvBase + INT#7] OR WORD#16#4000;
    END_IF;
// b15 BKRL／Control.BrakeRelease：TRUEはブレーキ強制解除。通常FALSE。縦軸では落下等の危険がある。
    IF RCON2_OUT[ConvAxisIndex].Control.BrakeRelease THEN
        RCON2_TxWord[ConvBase + INT#7] := RCON2_TxWord[ConvBase + INT#7] OR WORD#16#8000;
    END_IF;
END_FOR;

// 論理ワードから実際に送るUINTへ。INと同じ1ワード内のバイト交換を適用します。
FOR ConvWordIndex := INT#0 TO INT#47 DO
    ConvWord := RCON2_TxWord[ConvWordIndex];
    IF RCON2_SwapBytes THEN
        ConvWord := Swap(ConvWord);
    END_IF;
    RCON2_TxUInt[ConvWordIndex] := WORD_TO_UINT(ConvWord);
END_FOR;
(* Rung 458: 実I/O書込み（許可OFF=前値保持） *)
// 【RCON2／Node5／5軸】直接数値指定の通信変換。加速と減速は共通値です。
// 前提：全軸が直接数値指定、直動軸、共通8ワード＋軸番号順に各8ワード。実機の設定は別途照合。
// OUTはPLC→RCONの指令、INはRCON→PLCの現在値・状態。名前はPLCから見た方向です。
// 構造体は人が扱いやすい箱、Eで始まる変数はI/Oマップに割付済みの通信の出入口です。
// このSTは変換と許可付き代入までです。自動運転、通信正常判定、安全停止、開始受付の管理は含みません。
// Sysmacでの全体再ビルドと実機照合は未実施です。このファイルだけで実機へ転送しないでください。
// 【③ 確認・許可がそろったときだけ、実際のI/O出力変数へ書く】
// 初期状態はWriteEnable／LayoutConfirmed／ByteOrderConfirmed／CommOKがすべてFALSEです。
// これらを機械条件の確認なしに一括TRUEにしてはいけません。CommOKとMotionPermitは未作成です。
// FALSEのときは出力を更新しないだけ。前のStartやServoOnが残り得ます。停止指令ではありません。
// 安全停止・異常停止は別の設計です。書込み許可をOFFにすることを非常停止の代わりにしないでください。
// このSTだけでは動作開始しません。DSTR保持10ms以上、PEND OFF受付→DSTR OFF→PEND ON完了を管理する処理が必要です。
// GwWritten/AxisWrittenは「PLC変数へ代入した」印。通信成功・RCONの受付・移動完了を意味しません。
// 同じE始まりの出力変数を別のラダー/STから書くと、後から書いた値が優先します。出力担当を重複させないでください。

RCON2_GwWritten := FALSE;
FOR ConvAxisIndex := INT#1 TO INT#5 DO
    RCON2_AxisWritten[ConvAxisIndex] := FALSE;
END_FOR;

IF RCON2_WriteEnable AND RCON2_LayoutConfirmed AND RCON2_ByteOrderConfirmed AND RCON2_CommOK THEN
// 共通指令はMON/RTEのみ。最初のRUN応答に必要なため、軸DataValidとは別にGwApplyで許可します。
    IF RCON2_GwApply THEN
        E005_Out_OUT00_2003_01_1 := RCON2_TxUInt[0];
        RCON2_GwWritten := TRUE;
    END_IF;

// 1軸目＝実機軸No.0。OUT08～OUT15の8ワードをまとめて代入。
// AxisApply=この軸の更新許可、EncodeOK=変換OK、DataValid=入力情報の条件確認、MotionPermit=機械側の運転許可。
// 途中1ワードだけではなく、位置・幅・速度・加減速・押付け・制御を一組として渡します。
    IF RCON2_AxisApply[1] AND RCON2_EncodeOK[1] AND RCON2_IN[1].DataValid
       AND RCON2_MotionPermit[1] THEN
        E005_Out_OUT08_2003_09_1 := RCON2_TxUInt[8];
        E005_Out_OUT09_2003_0A_1 := RCON2_TxUInt[9];
        E005_Out_OUT10_2003_0B_1 := RCON2_TxUInt[10];
        E005_Out_OUT11_2003_0C_1 := RCON2_TxUInt[11];
        E005_Out_OUT12_2003_0D_1 := RCON2_TxUInt[12];
        E005_Out_OUT13_2003_0E_1 := RCON2_TxUInt[13];
        E005_Out_OUT14_2003_0F_1 := RCON2_TxUInt[14];
        E005_Out_OUT15_2003_10_1 := RCON2_TxUInt[15];
        RCON2_AxisWritten[1] := TRUE;
    END_IF;

// 2軸目＝実機軸No.1。OUT16～OUT23の8ワードをまとめて代入。
// AxisApply=この軸の更新許可、EncodeOK=変換OK、DataValid=入力情報の条件確認、MotionPermit=機械側の運転許可。
// 途中1ワードだけではなく、位置・幅・速度・加減速・押付け・制御を一組として渡します。
    IF RCON2_AxisApply[2] AND RCON2_EncodeOK[2] AND RCON2_IN[2].DataValid
       AND RCON2_MotionPermit[2] THEN
        E005_Out_OUT16_2003_11_1 := RCON2_TxUInt[16];
        E005_Out_OUT17_2003_12_1 := RCON2_TxUInt[17];
        E005_Out_OUT18_2003_13_1 := RCON2_TxUInt[18];
        E005_Out_OUT19_2003_14_1 := RCON2_TxUInt[19];
        E005_Out_OUT20_2003_15_1 := RCON2_TxUInt[20];
        E005_Out_OUT21_2003_16_1 := RCON2_TxUInt[21];
        E005_Out_OUT22_2003_17_1 := RCON2_TxUInt[22];
        E005_Out_OUT23_2003_18_1 := RCON2_TxUInt[23];
        RCON2_AxisWritten[2] := TRUE;
    END_IF;

// 3軸目＝実機軸No.2。OUT24～OUT31の8ワードをまとめて代入。
// AxisApply=この軸の更新許可、EncodeOK=変換OK、DataValid=入力情報の条件確認、MotionPermit=機械側の運転許可。
// 途中1ワードだけではなく、位置・幅・速度・加減速・押付け・制御を一組として渡します。
    IF RCON2_AxisApply[3] AND RCON2_EncodeOK[3] AND RCON2_IN[3].DataValid
       AND RCON2_MotionPermit[3] THEN
        E005_Out_OUT24_2003_19_1 := RCON2_TxUInt[24];
        E005_Out_OUT25_2003_1A_1 := RCON2_TxUInt[25];
        E005_Out_OUT26_2003_1B_1 := RCON2_TxUInt[26];
        E005_Out_OUT27_2003_1C_1 := RCON2_TxUInt[27];
        E005_Out_OUT28_2003_1D_1 := RCON2_TxUInt[28];
        E005_Out_OUT29_2003_1E_1 := RCON2_TxUInt[29];
        E005_Out_OUT30_2003_1F_1 := RCON2_TxUInt[30];
        E005_Out_OUT31_2003_20_1 := RCON2_TxUInt[31];
        RCON2_AxisWritten[3] := TRUE;
    END_IF;

// 4軸目＝実機軸No.3。OUT32～OUT39の8ワードをまとめて代入。
// AxisApply=この軸の更新許可、EncodeOK=変換OK、DataValid=入力情報の条件確認、MotionPermit=機械側の運転許可。
// 途中1ワードだけではなく、位置・幅・速度・加減速・押付け・制御を一組として渡します。
    IF RCON2_AxisApply[4] AND RCON2_EncodeOK[4] AND RCON2_IN[4].DataValid
       AND RCON2_MotionPermit[4] THEN
        E005_Out_OUT32_2003_21_1 := RCON2_TxUInt[32];
        E005_Out_OUT33_2003_22_1 := RCON2_TxUInt[33];
        E005_Out_OUT34_2003_23_1 := RCON2_TxUInt[34];
        E005_Out_OUT35_2003_24_1 := RCON2_TxUInt[35];
        E005_Out_OUT36_2003_25_1 := RCON2_TxUInt[36];
        E005_Out_OUT37_2003_26_1 := RCON2_TxUInt[37];
        E005_Out_OUT38_2003_27_1 := RCON2_TxUInt[38];
        E005_Out_OUT39_2003_28_1 := RCON2_TxUInt[39];
        RCON2_AxisWritten[4] := TRUE;
    END_IF;

// 5軸目＝実機軸No.4。OUT40～OUT47の8ワードをまとめて代入。
// AxisApply=この軸の更新許可、EncodeOK=変換OK、DataValid=入力情報の条件確認、MotionPermit=機械側の運転許可。
// 途中1ワードだけではなく、位置・幅・速度・加減速・押付け・制御を一組として渡します。
    IF RCON2_AxisApply[5] AND RCON2_EncodeOK[5] AND RCON2_IN[5].DataValid
       AND RCON2_MotionPermit[5] THEN
        E005_Out_OUT40_2003_29_1 := RCON2_TxUInt[40];
        E005_Out_OUT41_2003_2A_1 := RCON2_TxUInt[41];
        E005_Out_OUT42_2003_2B_1 := RCON2_TxUInt[42];
        E005_Out_OUT43_2003_2C_1 := RCON2_TxUInt[43];
        E005_Out_OUT44_2003_2D_1 := RCON2_TxUInt[44];
        E005_Out_OUT45_2003_2E_1 := RCON2_TxUInt[45];
        E005_Out_OUT46_2003_2F_1 := RCON2_TxUInt[46];
        E005_Out_OUT47_2003_30_1 := RCON2_TxUInt[47];
        RCON2_AxisWritten[5] := TRUE;
    END_IF;
END_IF;
// OUT01～07、OUT48～55は、このSTからは一切書き換えません。
// 現在の実機設定・別処理の用途が未確認なので、余剰領域を勝手にゼロクリアしません。

(* Section DLEP1_GT2: ladder, written here as Structured Text *)

